Universal Robots URScript: test_fourth_drawing_8_m18.script

def Machining4():
  # Default parameters:
  global speed_ms = 0.3
  global speed_rads = 0.75
  global accel_mss = 3
  global accel_radss = 1.2
  global blend_radius_m = 0.001

  # Add subprograms here
  # Start of main program
  # Program generated by RoboDK v5.6.5 for UR10e on 02/02/2024 17:39:49
  # Using nominal kinematics.
  blend_radius_m = 0.001
  speed_ms = 1.000
  # set_reference(p[0.348734, -0.005000, -0.017586, 0.000000, 0.000000, 0.000000])
  set_tcp(p[0.000000, 0.000000, 0.252000, 0.000000, 0.000000, 0.000000])
  # Show Tool
  movej([0.508484, -0.952512, -2.535391, -1.224486, 1.570796, 2.079280],accel_radss,speed_rads,0,blend_radius_m)
  movel([0.508484, -0.952512, -2.535391, -1.224486, 1.570796, 2.079280],accel_mss,speed_ms,0,blend_radius_m)
  # Splitting Linear movement in 6 (instruction 7: MoveL 3)
  movel([0.508484, -0.969998, -2.560672, -1.181720, 1.570796, 2.079280],accel_mss,speed_ms,0,blend_radius_m)
  movel([0.508484, -0.990214, -2.585461, -1.136714, 1.570796, 2.079280],accel_mss,speed_ms,0,blend_radius_m)
  movel([0.508484, -1.013449, -2.609714, -1.089227, 1.570796, 2.079280],accel_mss,speed_ms,0,blend_radius_m)
  movel([0.508484, -1.040019, -2.633377, -1.038993, 1.570796, 2.079280],accel_mss,speed_ms,0,blend_radius_m)
  movel([0.508484, -1.070270, -2.656387, -0.985731, 1.570796, 2.079280],accel_mss,speed_ms,0,blend_radius_m)
  movel([0.508484, -1.104577, -2.678669, -0.929143, 1.570796, 2.079280],accel_mss,speed_ms,0,blend_radius_m)
  movel([0.508484, -1.104577, -2.678669, -0.929143, 1.570796, 2.079280],accel_mss,speed_ms,0,blend_radius_m)
  speed_ms = 1.000
  movel([0.508484, -1.104577, -2.678669, -0.929143, 1.570796, 2.079280],accel_mss,speed_ms,0,blend_radius_m)
  movel([0.508484, -1.104577, -2.678669, -0.929143, 1.570796, 2.079280],accel_mss,speed_ms,0,blend_radius_m)
  movel([0.508484, -1.104577, -2.678669, -0.929143, 1.570796, 2.079280],accel_mss,speed_ms,0,blend_radius_m)
  speed_ms = 0.005
  movel([0.508484, -1.063908, -2.651841, -0.996640, 1.570796, 2.079280],accel_mss,speed_ms,0,blend_radius_m)
  speed_ms = 1.000
  movel([0.508484, -1.104577, -2.678669, -0.929143, 1.570796, 2.079280],accel_mss,speed_ms,0,blend_radius_m)
  speed_ms = 0.040
  movel([0.508484, -1.104577, -2.678669, -0.929143, 1.570796, 2.079280],accel_mss,speed_ms,0,blend_radius_m)
  speed_ms = 1.000
  movel([0.508484, -1.104577, -2.678669, -0.929143, 1.570796, 2.079280],accel_mss,speed_ms,0,blend_radius_m)
  # Splitting Linear movement in 8 (instruction 21: MoveL 12)
  movel([0.516357, -1.145060, -2.661765, -0.905563, 1.570796, 2.087153],accel_mss,speed_ms,0,blend_radius_m)
  movel([0.523521, -1.183921, -2.644010, -0.884457, 1.570796, 2.094317],accel_mss,speed_ms,0,blend_radius_m)
  movel([0.530064, -1.221217, -2.625467, -0.865705, 1.570796, 2.100861],accel_mss,speed_ms,0,blend_radius_m)
  movel([0.536061, -1.257021, -2.606194, -0.849174, 1.570796, 2.106857],accel_mss,speed_ms,0,blend_radius_m)
  movel([0.541574, -1.291418, -2.586246, -0.834725, 1.570796, 2.112371],accel_mss,speed_ms,0,blend_radius_m)
  movel([0.546659, -1.324498, -2.565672, -0.822220, 1.570796, 2.117455],accel_mss,speed_ms,0,blend_radius_m)
  movel([0.551360, -1.356351, -2.544515, -0.811522, 1.570796, 2.122157],accel_mss,speed_ms,0,blend_radius_m)
  movel([0.555720, -1.387070, -2.522816, -0.802503, 1.570796, 2.126517],accel_mss,speed_ms,0,blend_radius_m)
  speed_ms = 0.005
  movel([0.555720, -1.427952, -2.542321, -0.742116, 1.570796, 2.126517],accel_mss,speed_ms,0,blend_radius_m)
  speed_ms = 0.025
  movel([0.551886, -1.431799, -2.539331, -0.741259, 1.570796, 2.122682],accel_mss,speed_ms,0,blend_radius_m)
  movel([0.549891, -1.433665, -2.537873, -0.740851, 1.570796, 2.120688],accel_mss,speed_ms,0,blend_radius_m)
  movel([0.547837, -1.435468, -2.536459, -0.740462, 1.570796, 2.118634],accel_mss,speed_ms,0,blend_radius_m)
  movel([0.545720, -1.437189, -2.535105, -0.740095, 1.570796, 2.116517],accel_mss,speed_ms,0,blend_radius_m)
  movel([0.543536, -1.438810, -2.533826, -0.739753, 1.570796, 2.114332],accel_mss,speed_ms,0,blend_radius_m)
  movel([0.541277, -1.440313, -2.532636, -0.739441, 1.570796, 2.112073],accel_mss,speed_ms,0,blend_radius_m)
  movel([0.538938, -1.441676, -2.531553, -0.739160, 1.570796, 2.109734],accel_mss,speed_ms,0,blend_radius_m)
  movel([0.539897, -1.440992, -2.532097, -0.739300, 1.570796, 2.110693],accel_mss,speed_ms,0,blend_radius_m)
  movel([0.540974, -1.439974, -2.532904, -0.739511, 1.570796, 2.111771],accel_mss,speed_ms,0,blend_radius_m)
  movel([0.541871, -1.438872, -2.533777, -0.739741, 1.570796, 2.112668],accel_mss,speed_ms,0,blend_radius_m)
  movel([0.542155, -1.438369, -2.534174, -0.739846, 1.570796, 2.112951],accel_mss,speed_ms,0,blend_radius_m)
  movel([0.542280, -1.437941, -2.534512, -0.739936, 1.570796, 2.113076],accel_mss,speed_ms,0,blend_radius_m)
  movel([0.542211, -1.437608, -2.534775, -0.740006, 1.570796, 2.113008],accel_mss,speed_ms,0,blend_radius_m)
  movel([0.541951, -1.437454, -2.534896, -0.740039, 1.570796, 2.112747],accel_mss,speed_ms,0,blend_radius_m)
  movel([0.541528, -1.437461, -2.534891, -0.740037, 1.570796, 2.112324],accel_mss,speed_ms,0,blend_radius_m)
  movel([0.540960, -1.437607, -2.534776, -0.740007, 1.570796, 2.111756],accel_mss,speed_ms,0,blend_radius_m)
  movel([0.539505, -1.438234, -2.534280, -0.739874, 1.570796, 2.110301],accel_mss,speed_ms,0,blend_radius_m)
  movel([0.537786, -1.439172, -2.533539, -0.739678, 1.570796, 2.108582],accel_mss,speed_ms,0,blend_radius_m)
  movel([0.534336, -1.441332, -2.531826, -0.739230, 1.570796, 2.105133],accel_mss,speed_ms,0,blend_radius_m)
  movel([0.532176, -1.442774, -2.530679, -0.738936, 1.570796, 2.102972],accel_mss,speed_ms,0,blend_radius_m)
  movel([0.529059, -1.444697, -2.529144, -0.738548, 1.570796, 2.099855],accel_mss,speed_ms,0,blend_radius_m)
  movel([0.527463, -1.445498, -2.528503, -0.738388, 1.570796, 2.098260],accel_mss,speed_ms,0,blend_radius_m)
  movel([0.525843, -1.446095, -2.528025, -0.738269, 1.570796, 2.096640],accel_mss,speed_ms,0,blend_radius_m)
  movel([0.526257, -1.445821, -2.528245, -0.738324, 1.570796, 2.097053],accel_mss,speed_ms,0,blend_radius_m)
  movel([0.526732, -1.445268, -2.528687, -0.738434, 1.570796, 2.097529],accel_mss,speed_ms,0,blend_radius_m)
  movel([0.527721, -1.443665, -2.529968, -0.738755, 1.570796, 2.098517],accel_mss,speed_ms,0,blend_radius_m)
  movel([0.528500, -1.441980, -2.531312, -0.739098, 1.570796, 2.099296],accel_mss,speed_ms,0,blend_radius_m)
  movel([0.528712, -1.441319, -2.531837, -0.739233, 1.570796, 2.099508],accel_mss,speed_ms,0,blend_radius_m)
  movel([0.528754, -1.440900, -2.532170, -0.739319, 1.570796, 2.099550],accel_mss,speed_ms,0,blend_radius_m)
  movel([0.528518, -1.440358, -2.532599, -0.739431, 1.570796, 2.099315],accel_mss,speed_ms,0,blend_radius_m)
  movel([0.528131, -1.440101, -2.532804, -0.739485, 1.570796, 2.098927],accel_mss,speed_ms,0,blend_radius_m)
  movel([0.527622, -1.440071, -2.532827, -0.739491, 1.570796, 2.098419],accel_mss,speed_ms,0,blend_radius_m)
  movel([0.527024, -1.440220, -2.532709, -0.739460, 1.570796, 2.097821],accel_mss,speed_ms,0,blend_radius_m)
  movel([0.525708, -1.440829, -2.532226, -0.739334, 1.570796, 2.096504],accel_mss,speed_ms,0,blend_radius_m)
  movel([0.524451, -1.441503, -2.531691, -0.739195, 1.570796, 2.095247],accel_mss,speed_ms,0,blend_radius_m)
  movel([0.522478, -1.442423, -2.530959, -0.739007, 1.570796, 2.093274],accel_mss,speed_ms,0,blend_radius_m)
  movel([0.520576, -1.443144, -2.530385, -0.738861, 1.570796, 2.091372],accel_mss,speed_ms,0,blend_radius_m)
  movel([0.518692, -1.443593, -2.530026, -0.738770, 1.570796, 2.089489],accel_mss,speed_ms,0,blend_radius_m)
  movel([0.516787, -1.443689, -2.529949, -0.738750, 1.570796, 2.087583],accel_mss,speed_ms,0,blend_radius_m)
  movel([0.518245, -1.442894, -2.530584, -0.738911, 1.570796, 2.089042],accel_mss,speed_ms,0,blend_radius_m)
  movel([0.519593, -1.441927, -2.531353, -0.739108, 1.570796, 2.090389],accel_mss,speed_ms,0,blend_radius_m)
  movel([0.520169, -1.441329, -2.531829, -0.739231, 1.570796, 2.090965],accel_mss,speed_ms,0,blend_radius_m)
  movel([0.520610, -1.440680, -2.532344, -0.739365, 1.570796, 2.091406],accel_mss,speed_ms,0,blend_radius_m)
  movel([0.520870, -1.440025, -2.532863, -0.739500, 1.570796, 2.091666],accel_mss,speed_ms,0,blend_radius_m)
  movel([0.520888, -1.439417, -2.533345, -0.739627, 1.570796, 2.091684],accel_mss,speed_ms,0,blend_radius_m)
  movel([0.520543, -1.438832, -2.533808, -0.739749, 1.570796, 2.091340],accel_mss,speed_ms,0,blend_radius_m)
  movel([0.519903, -1.438483, -2.534084, -0.739822, 1.570796, 2.090700],accel_mss,speed_ms,0,blend_radius_m)
  movel([0.519080, -1.438310, -2.534221, -0.739858, 1.570796, 2.089876],accel_mss,speed_ms,0,blend_radius_m)
  movel([0.518194, -1.438247, -2.534271, -0.739872, 1.570796, 2.088990],accel_mss,speed_ms,0,blend_radius_m)
  speed_ms = 0.005
  movel([0.518194, -1.429866, -2.530530, -0.751993, 1.570796, 2.088990],accel_mss,speed_ms,0,blend_radius_m)
  speed_ms = 0.040
  movel([0.510141, -1.449455, -2.514970, -0.747963, 1.570796, 2.080938],accel_mss,speed_ms,0,blend_radius_m)
  speed_ms = 0.005
  movel([0.510141, -1.457684, -2.518629, -0.736076, 1.570796, 2.080938],accel_mss,speed_ms,0,blend_radius_m)
  speed_ms = 0.025
  movel([0.511091, -1.456693, -2.519440, -0.736256, 1.570796, 2.081888],accel_mss,speed_ms,0,blend_radius_m)
  movel([0.512141, -1.455770, -2.520195, -0.736424, 1.570796, 2.082937],accel_mss,speed_ms,0,blend_radius_m)
  movel([0.513267, -1.454927, -2.520883, -0.736579, 1.570796, 2.084063],accel_mss,speed_ms,0,blend_radius_m)
  movel([0.514457, -1.454175, -2.521496, -0.736718, 1.570796, 2.085253],accel_mss,speed_ms,0,blend_radius_m)
  movel([0.515692, -1.453521, -2.522028, -0.736840, 1.570796, 2.086488],accel_mss,speed_ms,0,blend_radius_m)
  movel([0.516954, -1.452980, -2.522467, -0.736941, 1.570796, 2.087750],accel_mss,speed_ms,0,blend_radius_m)
  movel([0.518224, -1.452560, -2.522808, -0.737020, 1.570796, 2.089020],accel_mss,speed_ms,0,blend_radius_m)
  movel([0.519487, -1.452271, -2.523043, -0.737075, 1.570796, 2.090284],accel_mss,speed_ms,0,blend_radius_m)
  movel([0.521308, -1.452078, -2.523200, -0.737111, 1.570796, 2.092104],accel_mss,speed_ms,0,blend_radius_m)
  movel([0.522944, -1.452159, -2.523134, -0.737096, 1.570796, 2.093740],accel_mss,speed_ms,0,blend_radius_m)
  movel([0.524404, -1.452488, -2.522867, -0.737034, 1.570796, 2.095200],accel_mss,speed_ms,0,blend_radius_m)
  movel([0.525694, -1.453041, -2.522418, -0.736930, 1.570796, 2.096491],accel_mss,speed_ms,0,blend_radius_m)
  movel([0.526823, -1.453792, -2.521807, -0.736790, 1.570796, 2.097619],accel_mss,speed_ms,0,blend_radius_m)
  movel([0.527798, -1.454719, -2.521052, -0.736618, 1.570796, 2.098594],accel_mss,speed_ms,0,blend_radius_m)
  movel([0.528624, -1.455797, -2.520173, -0.736419, 1.570796, 2.099421],accel_mss,speed_ms,0,blend_radius_m)
  movel([0.529313, -1.457000, -2.519189, -0.736200, 1.570796, 2.100109],accel_mss,speed_ms,0,blend_radius_m)
  movel([0.529870, -1.458305, -2.518119, -0.735965, 1.570796, 2.100667],accel_mss,speed_ms,0,blend_radius_m)
  movel([0.530307, -1.459689, -2.516982, -0.735718, 1.570796, 2.101103],accel_mss,speed_ms,0,blend_radius_m)
  movel([0.530848, -1.462592, -2.514587, -0.735210, 1.570796, 2.101644],accel_mss,speed_ms,0,blend_radius_m)
  movel([0.531006, -1.465517, -2.512160, -0.734712, 1.570796, 2.101803],accel_mss,speed_ms,0,blend_radius_m)
  movel([0.530842, -1.468282, -2.509854, -0.734253, 1.570796, 2.101639],accel_mss,speed_ms,0,blend_radius_m)
  movel([0.530390, -1.471193, -2.507413, -0.733783, 1.570796, 2.101186],accel_mss,speed_ms,0,blend_radius_m)
  movel([0.529720, -1.474131, -2.504936, -0.733322, 1.570796, 2.100516],accel_mss,speed_ms,0,blend_radius_m)
  movel([0.528861, -1.477086, -2.502431, -0.732872, 1.570796, 2.099658],accel_mss,speed_ms,0,blend_radius_m)
  movel([0.527841, -1.480049, -2.499906, -0.732435, 1.570796, 2.098637],accel_mss,speed_ms,0,blend_radius_m)
  movel([0.526687, -1.483008, -2.497369, -0.732012, 1.570796, 2.097483],accel_mss,speed_ms,0,blend_radius_m)
  movel([0.525429, -1.485956, -2.494829, -0.731604, 1.570796, 2.096225],accel_mss,speed_ms,0,blend_radius_m)
  movel([0.522707, -1.491776, -2.489774, -0.730839, 1.570796, 2.093504],accel_mss,speed_ms,0,blend_radius_m)
  movel([0.520789, -1.495817, -2.486233, -0.730340, 1.570796, 2.091586],accel_mss,speed_ms,0,blend_radius_m)
  movel([0.519999, -1.497823, -2.484465, -0.730101, 1.570796, 2.090795],accel_mss,speed_ms,0,blend_radius_m)
  movel([0.519432, -1.499808, -2.482709, -0.729872, 1.570796, 2.090228],accel_mss,speed_ms,0,blend_radius_m)
  movel([0.519026, -1.502378, -2.480427, -0.729584, 1.570796, 2.089822],accel_mss,speed_ms,0,blend_radius_m)
  movel([0.518624, -1.504952, -2.478131, -0.729306, 1.570796, 2.089420],accel_mss,speed_ms,0,blend_radius_m)
  movel([0.518292, -1.506214, -2.477001, -0.729174, 1.570796, 2.089088],accel_mss,speed_ms,0,blend_radius_m)
  movel([0.517800, -1.507448, -2.475895, -0.729047, 1.570796, 2.088596],accel_mss,speed_ms,0,blend_radius_m)
  movel([0.517098, -1.508640, -2.474823, -0.728926, 1.570796, 2.087894],accel_mss,speed_ms,0,blend_radius_m)
  movel([0.516134, -1.509785, -2.473791, -0.728813, 1.570796, 2.086930],accel_mss,speed_ms,0,blend_radius_m)
  movel([0.518755, -1.507097, -2.476210, -0.729083, 1.570796, 2.089552],accel_mss,speed_ms,0,blend_radius_m)
  movel([0.521247, -1.504345, -2.478673, -0.729371, 1.570796, 2.092043],accel_mss,speed_ms,0,blend_radius_m)
  movel([0.526020, -1.498683, -2.483705, -0.730001, 1.570796, 2.096816],accel_mss,speed_ms,0,blend_radius_m)
  movel([0.528599, -1.495468, -2.486539, -0.730382, 1.570796, 2.099395],accel_mss,speed_ms,0,blend_radius_m)
  movel([0.531106, -1.492207, -2.489397, -0.730784, 1.570796, 2.101903],accel_mss,speed_ms,0,blend_radius_m)
  movel([0.535966, -1.485569, -2.495163, -0.731657, 1.570796, 2.106762],accel_mss,speed_ms,0,blend_radius_m)
  movel([0.540563, -1.478943, -2.500850, -0.732596, 1.570796, 2.111359],accel_mss,speed_ms,0,blend_radius_m)
  movel([0.542732, -1.475555, -2.503731, -0.733104, 1.570796, 2.113528],accel_mss,speed_ms,0,blend_radius_m)
  movel([0.544723, -1.472142, -2.506614, -0.733633, 1.570796, 2.115519],accel_mss,speed_ms,0,blend_radius_m)
  movel([0.546112, -1.469422, -2.508900, -0.734068, 1.570796, 2.116908],accel_mss,speed_ms,0,blend_radius_m)
  movel([0.547394, -1.466668, -2.511201, -0.734519, 1.570796, 2.118190],accel_mss,speed_ms,0,blend_radius_m)
  movel([0.548701, -1.463889, -2.513512, -0.734988, 1.570796, 2.119497],accel_mss,speed_ms,0,blend_radius_m)
  movel([0.550164, -1.461093, -2.515825, -0.735471, 1.570796, 2.120961],accel_mss,speed_ms,0,blend_radius_m)
  movel([0.550637, -1.460364, -2.516426, -0.735599, 1.570796, 2.121434],accel_mss,speed_ms,0,blend_radius_m)
  movel([0.551236, -1.459675, -2.516993, -0.735720, 1.570796, 2.122032],accel_mss,speed_ms,0,blend_radius_m)
  movel([0.551916, -1.459170, -2.517409, -0.735810, 1.570796, 2.122713],accel_mss,speed_ms,0,blend_radius_m)
  movel([0.552279, -1.459029, -2.517525, -0.735835, 1.570796, 2.123075],accel_mss,speed_ms,0,blend_radius_m)
  movel([0.552650, -1.458984, -2.517562, -0.735843, 1.570796, 2.123447],accel_mss,speed_ms,0,blend_radius_m)
  movel([0.553094, -1.459095, -2.517470, -0.735823, 1.570796, 2.123890],accel_mss,speed_ms,0,blend_radius_m)
  movel([0.553450, -1.459322, -2.517284, -0.735783, 1.570796, 2.124247],accel_mss,speed_ms,0,blend_radius_m)
  movel([0.555162, -1.460824, -2.516047, -0.735518, 1.570796, 2.125958],accel_mss,speed_ms,0,blend_radius_m)
  movel([0.556530, -1.462499, -2.514664, -0.735226, 1.570796, 2.127326],accel_mss,speed_ms,0,blend_radius_m)
  movel([0.557585, -1.464326, -2.513150, -0.734913, 1.570796, 2.128381],accel_mss,speed_ms,0,blend_radius_m)
  movel([0.558352, -1.466294, -2.511513, -0.734582, 1.570796, 2.129148],accel_mss,speed_ms,0,blend_radius_m)
  movel([0.558858, -1.468380, -2.509772, -0.734237, 1.570796, 2.129655],accel_mss,speed_ms,0,blend_radius_m)
  movel([0.559133, -1.470569, -2.507937, -0.733883, 1.570796, 2.129930],accel_mss,speed_ms,0,blend_radius_m)
  movel([0.559203, -1.472844, -2.506022, -0.733522, 1.570796, 2.129999],accel_mss,speed_ms,0,blend_radius_m)
  movel([0.559091, -1.475191, -2.504039, -0.733159, 1.570796, 2.129888],accel_mss,speed_ms,0,blend_radius_m)
  movel([0.558827, -1.477592, -2.502001, -0.732796, 1.570796, 2.129624],accel_mss,speed_ms,0,blend_radius_m)
  movel([0.558438, -1.480032, -2.499920, -0.732437, 1.570796, 2.129235],accel_mss,speed_ms,0,blend_radius_m)
  movel([0.557386, -1.484964, -2.495685, -0.731739, 1.570796, 2.128183],accel_mss,speed_ms,0,blend_radius_m)
  movel([0.554892, -1.494646, -2.487262, -0.730482, 1.570796, 2.125689],accel_mss,speed_ms,0,blend_radius_m)
  movel([0.554588, -1.496145, -2.485944, -0.730300, 1.570796, 2.125384],accel_mss,speed_ms,0,blend_radius_m)
  movel([0.554575, -1.496851, -2.485322, -0.730216, 1.570796, 2.125371],accel_mss,speed_ms,0,blend_radius_m)
  movel([0.554722, -1.497492, -2.484757, -0.730140, 1.570796, 2.125519],accel_mss,speed_ms,0,blend_radius_m)
  movel([0.555275, -1.498243, -2.484094, -0.730052, 1.570796, 2.126071],accel_mss,speed_ms,0,blend_radius_m)
  movel([0.555655, -1.498482, -2.483883, -0.730024, 1.570796, 2.126451],accel_mss,speed_ms,0,blend_radius_m)
  movel([0.556095, -1.498637, -2.483746, -0.730006, 1.570796, 2.126891],accel_mss,speed_ms,0,blend_radius_m)
  movel([0.557113, -1.498726, -2.483667, -0.729996, 1.570796, 2.127910],accel_mss,speed_ms,0,blend_radius_m)
  movel([0.558266, -1.498560, -2.483813, -0.730015, 1.570796, 2.129063],accel_mss,speed_ms,0,blend_radius_m)
  movel([0.559484, -1.498195, -2.484136, -0.730058, 1.570796, 2.130280],accel_mss,speed_ms,0,blend_radius_m)
  movel([0.560700, -1.497680, -2.484591, -0.730118, 1.570796, 2.131496],accel_mss,speed_ms,0,blend_radius_m)
  movel([0.561849, -1.497066, -2.485132, -0.730190, 1.570796, 2.132646],accel_mss,speed_ms,0,blend_radius_m)
  movel([0.562859, -1.496403, -2.485717, -0.730269, 1.570796, 2.133656],accel_mss,speed_ms,0,blend_radius_m)
  movel([0.564501, -1.495161, -2.486809, -0.730419, 1.570796, 2.135297],accel_mss,speed_ms,0,blend_radius_m)
  movel([0.566103, -1.493854, -2.487956, -0.730579, 1.570796, 2.136900],accel_mss,speed_ms,0,blend_radius_m)
  movel([0.569169, -1.491072, -2.490389, -0.730929, 1.570796, 2.139965],accel_mss,speed_ms,0,blend_radius_m)
  movel([0.572027, -1.488119, -2.492957, -0.731313, 1.570796, 2.142824],accel_mss,speed_ms,0,blend_radius_m)
  movel([0.574646, -1.485054, -2.495608, -0.731727, 1.570796, 2.145443],accel_mss,speed_ms,0,blend_radius_m)
  movel([0.575591, -1.483880, -2.496620, -0.731890, 1.570796, 2.146387],accel_mss,speed_ms,0,blend_radius_m)
  movel([0.576618, -1.482762, -2.497581, -0.732046, 1.570796, 2.147414],accel_mss,speed_ms,0,blend_radius_m)
  movel([0.577188, -1.482268, -2.498005, -0.732116, 1.570796, 2.147985],accel_mss,speed_ms,0,blend_radius_m)
  movel([0.577814, -1.481835, -2.498377, -0.732178, 1.570796, 2.148610],accel_mss,speed_ms,0,blend_radius_m)
  movel([0.578503, -1.481482, -2.498679, -0.732228, 1.570796, 2.149299],accel_mss,speed_ms,0,blend_radius_m)
  movel([0.579266, -1.481229, -2.498896, -0.732264, 1.570796, 2.150062],accel_mss,speed_ms,0,blend_radius_m)
  movel([0.580251, -1.481159, -2.498956, -0.732274, 1.570796, 2.151047],accel_mss,speed_ms,0,blend_radius_m)
  movel([0.581073, -1.481422, -2.498731, -0.732237, 1.570796, 2.151869],accel_mss,speed_ms,0,blend_radius_m)
  movel([0.581707, -1.481932, -2.498293, -0.732164, 1.570796, 2.152503],accel_mss,speed_ms,0,blend_radius_m)
  movel([0.582136, -1.482605, -2.497715, -0.732068, 1.570796, 2.152933],accel_mss,speed_ms,0,blend_radius_m)
  movel([0.582578, -1.483885, -2.496615, -0.731889, 1.570796, 2.153374],accel_mss,speed_ms,0,blend_radius_m)
  movel([0.582850, -1.485265, -2.495426, -0.731698, 1.570796, 2.153646],accel_mss,speed_ms,0,blend_radius_m)
  movel([0.583065, -1.488131, -2.492947, -0.731312, 1.570796, 2.153861],accel_mss,speed_ms,0,blend_radius_m)
  movel([0.583037, -1.489513, -2.491746, -0.731130, 1.570796, 2.153834],accel_mss,speed_ms,0,blend_radius_m)
  movel([0.582882, -1.490891, -2.490546, -0.730952, 1.570796, 2.153679],accel_mss,speed_ms,0,blend_radius_m)
  movel([0.582611, -1.492261, -2.489350, -0.730778, 1.570796, 2.153407],accel_mss,speed_ms,0,blend_radius_m)
  movel([0.582227, -1.493625, -2.488157, -0.730607, 1.570796, 2.153023],accel_mss,speed_ms,0,blend_radius_m)
  movel([0.581738, -1.494980, -2.486969, -0.730441, 1.570796, 2.152535],accel_mss,speed_ms,0,blend_radius_m)
  movel([0.580473, -1.497665, -2.484604, -0.730120, 1.570796, 2.151270],accel_mss,speed_ms,0,blend_radius_m)
  movel([0.579710, -1.498992, -2.483432, -0.729965, 1.570796, 2.150506],accel_mss,speed_ms,0,blend_radius_m)
  movel([0.577960, -1.501613, -2.481108, -0.729668, 1.570796, 2.148756],accel_mss,speed_ms,0,blend_radius_m)
  movel([0.575952, -1.504185, -2.478816, -0.729388, 1.570796, 2.146749],accel_mss,speed_ms,0,blend_radius_m)
  movel([0.573737, -1.506705, -2.476561, -0.729123, 1.570796, 2.144533],accel_mss,speed_ms,0,blend_radius_m)
  movel([0.571371, -1.509163, -2.474352, -0.728874, 1.570796, 2.142167],accel_mss,speed_ms,0,blend_radius_m)
  movel([0.567732, -1.512631, -2.471218, -0.728540, 1.570796, 2.138528],accel_mss,speed_ms,0,blend_radius_m)
  movel([0.565824, -1.514296, -2.469707, -0.728386, 1.570796, 2.136621],accel_mss,speed_ms,0,blend_radius_m)
  movel([0.563854, -1.515893, -2.468253, -0.728243, 1.570796, 2.134651],accel_mss,speed_ms,0,blend_radius_m)
  movel([0.561822, -1.517401, -2.466876, -0.728112, 1.570796, 2.132618],accel_mss,speed_ms,0,blend_radius_m)
  movel([0.559727, -1.518806, -2.465590, -0.727992, 1.570796, 2.130523],accel_mss,speed_ms,0,blend_radius_m)
  movel([0.557561, -1.520091, -2.464412, -0.727886, 1.570796, 2.128357],accel_mss,speed_ms,0,blend_radius_m)
  movel([0.555327, -1.521236, -2.463359, -0.727794, 1.570796, 2.126124],accel_mss,speed_ms,0,blend_radius_m)
  movel([0.552124, -1.522621, -2.462084, -0.727685, 1.570796, 2.122920],accel_mss,speed_ms,0,blend_radius_m)
  movel([0.550419, -1.523230, -2.461521, -0.727638, 1.570796, 2.121215],accel_mss,speed_ms,0,blend_radius_m)
  movel([0.548705, -1.523722, -2.461067, -0.727600, 1.570796, 2.119502],accel_mss,speed_ms,0,blend_radius_m)
  movel([0.547032, -1.524050, -2.460764, -0.727575, 1.570796, 2.117828],accel_mss,speed_ms,0,blend_radius_m)
  movel([0.545444, -1.524166, -2.460656, -0.727567, 1.570796, 2.116240],accel_mss,speed_ms,0,blend_radius_m)
  movel([0.543989, -1.524022, -2.460790, -0.727577, 1.570796, 2.114785],accel_mss,speed_ms,0,blend_radius_m)
  movel([0.543326, -1.523839, -2.460959, -0.727591, 1.570796, 2.114122],accel_mss,speed_ms,0,blend_radius_m)
  movel([0.542715, -1.523572, -2.461206, -0.727611, 1.570796, 2.113512],accel_mss,speed_ms,0,blend_radius_m)
  movel([0.542106, -1.523172, -2.461575, -0.727642, 1.570796, 2.112902],accel_mss,speed_ms,0,blend_radius_m)
  movel([0.541607, -1.522687, -2.462022, -0.727679, 1.570796, 2.112403],accel_mss,speed_ms,0,blend_radius_m)
  movel([0.541207, -1.522126, -2.462540, -0.727723, 1.570796, 2.112004],accel_mss,speed_ms,0,blend_radius_m)
  movel([0.540902, -1.521496, -2.463120, -0.727773, 1.570796, 2.111698],accel_mss,speed_ms,0,blend_radius_m)
  movel([0.540535, -1.520068, -2.464433, -0.727888, 1.570796, 2.111331],accel_mss,speed_ms,0,blend_radius_m)
  movel([0.540444, -1.518473, -2.465896, -0.728020, 1.570796, 2.111240],accel_mss,speed_ms,0,blend_radius_m)
  movel([0.540559, -1.516785, -2.467439, -0.728165, 1.570796, 2.111355],accel_mss,speed_ms,0,blend_radius_m)
  movel([0.540816, -1.515077, -2.468996, -0.728316, 1.570796, 2.111612],accel_mss,speed_ms,0,blend_radius_m)
  movel([0.541487, -1.511892, -2.471888, -0.728610, 1.570796, 2.112284],accel_mss,speed_ms,0,blend_radius_m)
  movel([0.541819, -1.510404, -2.473232, -0.728752, 1.570796, 2.112615],accel_mss,speed_ms,0,blend_radius_m)
  movel([0.541998, -1.508958, -2.474537, -0.728895, 1.570796, 2.112794],accel_mss,speed_ms,0,blend_radius_m)
  movel([0.541952, -1.508290, -2.475137, -0.728961, 1.570796, 2.112748],accel_mss,speed_ms,0,blend_radius_m)
  movel([0.541774, -1.507681, -2.475685, -0.729023, 1.570796, 2.112571],accel_mss,speed_ms,0,blend_radius_m)
  movel([0.541434, -1.507148, -2.476163, -0.729077, 1.570796, 2.112230],accel_mss,speed_ms,0,blend_radius_m)
  movel([0.540901, -1.506706, -2.476560, -0.729123, 1.570796, 2.111697],accel_mss,speed_ms,0,blend_radius_m)
  movel([0.540999, -1.506837, -2.476443, -0.729109, 1.570796, 2.111796],accel_mss,speed_ms,0,blend_radius_m)
  movel([0.540993, -1.507039, -2.476261, -0.729088, 1.570796, 2.111789],accel_mss,speed_ms,0,blend_radius_m)
  movel([0.540687, -1.507637, -2.475725, -0.729027, 1.570796, 2.111483],accel_mss,speed_ms,0,blend_radius_m)
  movel([0.540031, -1.508460, -2.474985, -0.728944, 1.570796, 2.110827],accel_mss,speed_ms,0,blend_radius_m)
  movel([0.539081, -1.509472, -2.474073, -0.728844, 1.570796, 2.109877],accel_mss,speed_ms,0,blend_radius_m)
  movel([0.536506, -1.511911, -2.471870, -0.728608, 1.570796, 2.107302],accel_mss,speed_ms,0,blend_radius_m)
  movel([0.533377, -1.514652, -2.469383, -0.728354, 1.570796, 2.104174],accel_mss,speed_ms,0,blend_radius_m)
  movel([0.527088, -1.519857, -2.464627, -0.727905, 1.570796, 2.097884],accel_mss,speed_ms,0,blend_radius_m)
  movel([0.523408, -1.522733, -2.461980, -0.727676, 1.570796, 2.094204],accel_mss,speed_ms,0,blend_radius_m)
  movel([0.519372, -1.525494, -2.459426, -0.727468, 1.570796, 2.090168],accel_mss,speed_ms,0,blend_radius_m)
  movel([0.515337, -1.528147, -2.456962, -0.727280, 1.570796, 2.086134],accel_mss,speed_ms,0,blend_radius_m)
  movel([0.511276, -1.530728, -2.454553, -0.727108, 1.570796, 2.082072],accel_mss,speed_ms,0,blend_radius_m)
  movel([0.503302, -1.535575, -2.450000, -0.726814, 1.570796, 2.074098],accel_mss,speed_ms,0,blend_radius_m)
  movel([0.499392, -1.537721, -2.447972, -0.726695, 1.570796, 2.070188],accel_mss,speed_ms,0,blend_radius_m)
  movel([0.497416, -1.538674, -2.447070, -0.726645, 1.570796, 2.068213],accel_mss,speed_ms,0,blend_radius_m)
  movel([0.495430, -1.539517, -2.446269, -0.726602, 1.570796, 2.066226],accel_mss,speed_ms,0,blend_radius_m)
  movel([0.493429, -1.540226, -2.445596, -0.726567, 1.570796, 2.064225],accel_mss,speed_ms,0,blend_radius_m)
  movel([0.491417, -1.540779, -2.445070, -0.726540, 1.570796, 2.062214],accel_mss,speed_ms,0,blend_radius_m)
  movel([0.493294, -1.537726, -2.447968, -0.726695, 1.570796, 2.064090],accel_mss,speed_ms,0,blend_radius_m)
  movel([0.493731, -1.536801, -2.448843, -0.726745, 1.570796, 2.064527],accel_mss,speed_ms,0,blend_radius_m)
  movel([0.493771, -1.536384, -2.449237, -0.726768, 1.570796, 2.064567],accel_mss,speed_ms,0,blend_radius_m)
  movel([0.493597, -1.536066, -2.449537, -0.726786, 1.570796, 2.064394],accel_mss,speed_ms,0,blend_radius_m)
  movel([0.493297, -1.535935, -2.449661, -0.726793, 1.570796, 2.064093],accel_mss,speed_ms,0,blend_radius_m)
  movel([0.492915, -1.535922, -2.449673, -0.726794, 1.570796, 2.063711],accel_mss,speed_ms,0,blend_radius_m)
  movel([0.490914, -1.536231, -2.449382, -0.726777, 1.570796, 2.061711],accel_mss,speed_ms,0,blend_radius_m)
  movel([0.489818, -1.536232, -2.449381, -0.726777, 1.570796, 2.060615],accel_mss,speed_ms,0,blend_radius_m)
  movel([0.488797, -1.536075, -2.449529, -0.726785, 1.570796, 2.059594],accel_mss,speed_ms,0,blend_radius_m)
  movel([0.487879, -1.535763, -2.449823, -0.726803, 1.570796, 2.058675],accel_mss,speed_ms,0,blend_radius_m)
  movel([0.487648, -1.535578, -2.449998, -0.726813, 1.570796, 2.058445],accel_mss,speed_ms,0,blend_radius_m)
  movel([0.487677, -1.535333, -2.450228, -0.726827, 1.570796, 2.058473],accel_mss,speed_ms,0,blend_radius_m)
  movel([0.488374, -1.534524, -2.450991, -0.726874, 1.570796, 2.059170],accel_mss,speed_ms,0,blend_radius_m)
  movel([0.488495, -1.534216, -2.451281, -0.726892, 1.570796, 2.059291],accel_mss,speed_ms,0,blend_radius_m)
  movel([0.488458, -1.533935, -2.451545, -0.726909, 1.570796, 2.059254],accel_mss,speed_ms,0,blend_radius_m)
  movel([0.488296, -1.533709, -2.451758, -0.726922, 1.570796, 2.059092],accel_mss,speed_ms,0,blend_radius_m)
  movel([0.488039, -1.533564, -2.451894, -0.726931, 1.570796, 2.058835],accel_mss,speed_ms,0,blend_radius_m)
  movel([0.487372, -1.533509, -2.451945, -0.726934, 1.570796, 2.058169],accel_mss,speed_ms,0,blend_radius_m)
  movel([0.482012, -1.534472, -2.451040, -0.726877, 1.570796, 2.052809],accel_mss,speed_ms,0,blend_radius_m)
  movel([0.483729, -1.533917, -2.451562, -0.726910, 1.570796, 2.054525],accel_mss,speed_ms,0,blend_radius_m)
  movel([0.485480, -1.533241, -2.452198, -0.726951, 1.570796, 2.056276],accel_mss,speed_ms,0,blend_radius_m)
  movel([0.487243, -1.532463, -2.452928, -0.726998, 1.570796, 2.058040],accel_mss,speed_ms,0,blend_radius_m)
  movel([0.489007, -1.531599, -2.453738, -0.727052, 1.570796, 2.059803],accel_mss,speed_ms,0,blend_radius_m)
  movel([0.492467, -1.529679, -2.455534, -0.727177, 1.570796, 2.063264],accel_mss,speed_ms,0,blend_radius_m)
  movel([0.495725, -1.527617, -2.457455, -0.727317, 1.570796, 2.066521],accel_mss,speed_ms,0,blend_radius_m)
  movel([0.499158, -1.525260, -2.459643, -0.727485, 1.570796, 2.069954],accel_mss,speed_ms,0,blend_radius_m)
  movel([0.502533, -1.522773, -2.461943, -0.727673, 1.570796, 2.073330],accel_mss,speed_ms,0,blend_radius_m)
  movel([0.504170, -1.521467, -2.463147, -0.727775, 1.570796, 2.074966],accel_mss,speed_ms,0,blend_radius_m)
  movel([0.505759, -1.520115, -2.464390, -0.727884, 1.570796, 2.076556],accel_mss,speed_ms,0,blend_radius_m)
  movel([0.507286, -1.518712, -2.465677, -0.728000, 1.570796, 2.078082],accel_mss,speed_ms,0,blend_radius_m)
  movel([0.508742, -1.517249, -2.467015, -0.728125, 1.570796, 2.079538],accel_mss,speed_ms,0,blend_radius_m)
  movel([0.509588, -1.516300, -2.467881, -0.728207, 1.570796, 2.080384],accel_mss,speed_ms,0,blend_radius_m)
  movel([0.510366, -1.515308, -2.468786, -0.728295, 1.570796, 2.081163],accel_mss,speed_ms,0,blend_radius_m)
  movel([0.511731, -1.513219, -2.470684, -0.728485, 1.570796, 2.082527],accel_mss,speed_ms,0,blend_radius_m)
  movel([0.512844, -1.511031, -2.472666, -0.728692, 1.570796, 2.083641],accel_mss,speed_ms,0,blend_radius_m)
  movel([0.513716, -1.508789, -2.474689, -0.728912, 1.570796, 2.084513],accel_mss,speed_ms,0,blend_radius_m)
  movel([0.514362, -1.506538, -2.476711, -0.729140, 1.570796, 2.085158],accel_mss,speed_ms,0,blend_radius_m)
  movel([0.514791, -1.504328, -2.478688, -0.729372, 1.570796, 2.085588],accel_mss,speed_ms,0,blend_radius_m)
  movel([0.515013, -1.502206, -2.480580, -0.729603, 1.570796, 2.085809],accel_mss,speed_ms,0,blend_radius_m)
  movel([0.515040, -1.500220, -2.482344, -0.729825, 1.570796, 2.085836],accel_mss,speed_ms,0,blend_radius_m)
  movel([0.514833, -1.499178, -2.483268, -0.729944, 1.570796, 2.085629],accel_mss,speed_ms,0,blend_radius_m)
  movel([0.514328, -1.498388, -2.483965, -0.730035, 1.570796, 2.085125],accel_mss,speed_ms,0,blend_radius_m)
  movel([0.513576, -1.497861, -2.484431, -0.730097, 1.570796, 2.084372],accel_mss,speed_ms,0,blend_radius_m)
  movel([0.512626, -1.497606, -2.484656, -0.730127, 1.570796, 2.083422],accel_mss,speed_ms,0,blend_radius_m)
  movel([0.511527, -1.497627, -2.484638, -0.730124, 1.570796, 2.082323],accel_mss,speed_ms,0,blend_radius_m)
  movel([0.510328, -1.497933, -2.484368, -0.730088, 1.570796, 2.081125],accel_mss,speed_ms,0,blend_radius_m)
  movel([0.509087, -1.498529, -2.483841, -0.730019, 1.570796, 2.079883],accel_mss,speed_ms,0,blend_radius_m)
  movel([0.507849, -1.499420, -2.483053, -0.729916, 1.570796, 2.078646],accel_mss,speed_ms,0,blend_radius_m)
  movel([0.506057, -1.500901, -2.481740, -0.729748, 1.570796, 2.076853],accel_mss,speed_ms,0,blend_radius_m)
  movel([0.504215, -1.502308, -2.480490, -0.729592, 1.570796, 2.075011],accel_mss,speed_ms,0,blend_radius_m)
  movel([0.502327, -1.503615, -2.479325, -0.729449, 1.570796, 2.073123],accel_mss,speed_ms,0,blend_radius_m)
  movel([0.500388, -1.504800, -2.478267, -0.729322, 1.570796, 2.071184],accel_mss,speed_ms,0,blend_radius_m)
  movel([0.498404, -1.505837, -2.477339, -0.729213, 1.570796, 2.069200],accel_mss,speed_ms,0,blend_radius_m)
  movel([0.496371, -1.506704, -2.476562, -0.729123, 1.570796, 2.067167],accel_mss,speed_ms,0,blend_radius_m)
  movel([0.494289, -1.507378, -2.475957, -0.729054, 1.570796, 2.065085],accel_mss,speed_ms,0,blend_radius_m)
  movel([0.492160, -1.507833, -2.475548, -0.729008, 1.570796, 2.062956],accel_mss,speed_ms,0,blend_radius_m)
  movel([0.491077, -1.507930, -2.475462, -0.728998, 1.570796, 2.061873],accel_mss,speed_ms,0,blend_radius_m)
  movel([0.490044, -1.507891, -2.475496, -0.729002, 1.570796, 2.060840],accel_mss,speed_ms,0,blend_radius_m)
  movel([0.488081, -1.507580, -2.475776, -0.729033, 1.570796, 2.058877],accel_mss,speed_ms,0,blend_radius_m)
  movel([0.486632, -1.507175, -2.476139, -0.729075, 1.570796, 2.057428],accel_mss,speed_ms,0,blend_radius_m)
  movel([0.485361, -1.506589, -2.476665, -0.729135, 1.570796, 2.056158],accel_mss,speed_ms,0,blend_radius_m)
  movel([0.484262, -1.505838, -2.477338, -0.729213, 1.570796, 2.055058],accel_mss,speed_ms,0,blend_radius_m)
  movel([0.483321, -1.504938, -2.478144, -0.729308, 1.570796, 2.054117],accel_mss,speed_ms,0,blend_radius_m)
  movel([0.482527, -1.503906, -2.479066, -0.729418, 1.570796, 2.053323],accel_mss,speed_ms,0,blend_radius_m)
  movel([0.481869, -1.502756, -2.480091, -0.729542, 1.570796, 2.052665],accel_mss,speed_ms,0,blend_radius_m)
  movel([0.481342, -1.501504, -2.481204, -0.729680, 1.570796, 2.052138],accel_mss,speed_ms,0,blend_radius_m)
  movel([0.480931, -1.500169, -2.482389, -0.729831, 1.570796, 2.051727],accel_mss,speed_ms,0,blend_radius_m)
  movel([0.480626, -1.498766, -2.483631, -0.729991, 1.570796, 2.051422],accel_mss,speed_ms,0,blend_radius_m)
  movel([0.480420, -1.497308, -2.484919, -0.730162, 1.570796, 2.051216],accel_mss,speed_ms,0,blend_radius_m)
  movel([0.480258, -1.494306, -2.487560, -0.730523, 1.570796, 2.051054],accel_mss,speed_ms,0,blend_radius_m)
  movel([0.480362, -1.491291, -2.490197, -0.730901, 1.570796, 2.051158],accel_mss,speed_ms,0,blend_radius_m)
  movel([0.480649, -1.488405, -2.492708, -0.731275, 1.570796, 2.051445],accel_mss,speed_ms,0,blend_radius_m)
  movel([0.480991, -1.486173, -2.494642, -0.731574, 1.570796, 2.051788],accel_mss,speed_ms,0,blend_radius_m)
  movel([0.481470, -1.483852, -2.496643, -0.731893, 1.570796, 2.052266],accel_mss,speed_ms,0,blend_radius_m)
  movel([0.482087, -1.481456, -2.498701, -0.732232, 1.570796, 2.052883],accel_mss,speed_ms,0,blend_radius_m)
  movel([0.482851, -1.479008, -2.500794, -0.732587, 1.570796, 2.053648],accel_mss,speed_ms,0,blend_radius_m)
  movel([0.483763, -1.476523, -2.502909, -0.732957, 1.570796, 2.054560],accel_mss,speed_ms,0,blend_radius_m)
  movel([0.484830, -1.474022, -2.505028, -0.733339, 1.570796, 2.055627],accel_mss,speed_ms,0,blend_radius_m)
  movel([0.486057, -1.471525, -2.507134, -0.733730, 1.570796, 2.056854],accel_mss,speed_ms,0,blend_radius_m)
  movel([0.487449, -1.469050, -2.509211, -0.734128, 1.570796, 2.058245],accel_mss,speed_ms,0,blend_radius_m)
  movel([0.489008, -1.466616, -2.511245, -0.734528, 1.570796, 2.059805],accel_mss,speed_ms,0,blend_radius_m)
  movel([0.490739, -1.464248, -2.513215, -0.734927, 1.570796, 2.061535],accel_mss,speed_ms,0,blend_radius_m)
  movel([0.492647, -1.461961, -2.515109, -0.735320, 1.570796, 2.063443],accel_mss,speed_ms,0,blend_radius_m)
  movel([0.494736, -1.459780, -2.516907, -0.735702, 1.570796, 2.065532],accel_mss,speed_ms,0,blend_radius_m)
  movel([0.497007, -1.457726, -2.518594, -0.736069, 1.570796, 2.067803],accel_mss,speed_ms,0,blend_radius_m)
  movel([0.499467, -1.455820, -2.520154, -0.736415, 1.570796, 2.070264],accel_mss,speed_ms,0,blend_radius_m)
  movel([0.502114, -1.454087, -2.521567, -0.736735, 1.570796, 2.072911],accel_mss,speed_ms,0,blend_radius_m)
  movel([0.504952, -1.452548, -2.522818, -0.737023, 1.570796, 2.075748],accel_mss,speed_ms,0,blend_radius_m)
  movel([0.506085, -1.452062, -2.523213, -0.737114, 1.570796, 2.076882],accel_mss,speed_ms,0,blend_radius_m)
  movel([0.506646, -1.451910, -2.523336, -0.737143, 1.570796, 2.077442],accel_mss,speed_ms,0,blend_radius_m)
  movel([0.507180, -1.451865, -2.523372, -0.737151, 1.570796, 2.077976],accel_mss,speed_ms,0,blend_radius_m)
  movel([0.507850, -1.452048, -2.523224, -0.737117, 1.570796, 2.078646],accel_mss,speed_ms,0,blend_radius_m)
  movel([0.508305, -1.452476, -2.522877, -0.737036, 1.570796, 2.079101],accel_mss,speed_ms,0,blend_radius_m)
  movel([0.508559, -1.453073, -2.522392, -0.736924, 1.570796, 2.079355],accel_mss,speed_ms,0,blend_radius_m)
  movel([0.508624, -1.453762, -2.521832, -0.736795, 1.570796, 2.079421],accel_mss,speed_ms,0,blend_radius_m)
  movel([0.508371, -1.455391, -2.520505, -0.736494, 1.570796, 2.079167],accel_mss,speed_ms,0,blend_radius_m)
  movel([0.507807, -1.457086, -2.519119, -0.736184, 1.570796, 2.078604],accel_mss,speed_ms,0,blend_radius_m)
  movel([0.506383, -1.460472, -2.516337, -0.735580, 1.570796, 2.077180],accel_mss,speed_ms,0,blend_radius_m)
  movel([0.506259, -1.461115, -2.515807, -0.735467, 1.570796, 2.077056],accel_mss,speed_ms,0,blend_radius_m)
  movel([0.506393, -1.461311, -2.515645, -0.735433, 1.570796, 2.077189],accel_mss,speed_ms,0,blend_radius_m)
  movel([0.506705, -1.461409, -2.515565, -0.735416, 1.570796, 2.077502],accel_mss,speed_ms,0,blend_radius_m)
  movel([0.507835, -1.460385, -2.516409, -0.735595, 1.570796, 2.078631],accel_mss,speed_ms,0,blend_radius_m)
  movel([0.508922, -1.459289, -2.517311, -0.735789, 1.570796, 2.079718],accel_mss,speed_ms,0,blend_radius_m)
  movel([0.506690, -1.464208, -2.513247, -0.734933, 1.570796, 2.077486],accel_mss,speed_ms,0,blend_radius_m)
  movel([0.504647, -1.469094, -2.509174, -0.734121, 1.570796, 2.075443],accel_mss,speed_ms,0,blend_radius_m)
  movel([0.502794, -1.473940, -2.505097, -0.733352, 1.570796, 2.073591],accel_mss,speed_ms,0,blend_radius_m)
  movel([0.501130, -1.478747, -2.501017, -0.732625, 1.570796, 2.071926],accel_mss,speed_ms,0,blend_radius_m)
  movel([0.500482, -1.480827, -2.499240, -0.732322, 1.570796, 2.071279],accel_mss,speed_ms,0,blend_radius_m)
  movel([0.499986, -1.482980, -2.497394, -0.732016, 1.570796, 2.070782],accel_mss,speed_ms,0,blend_radius_m)
  movel([0.499855, -1.484030, -2.496490, -0.731869, 1.570796, 2.070651],accel_mss,speed_ms,0,blend_radius_m)
  movel([0.499835, -1.485034, -2.495625, -0.731730, 1.570796, 2.070632],accel_mss,speed_ms,0,blend_radius_m)
  movel([0.499953, -1.485969, -2.494818, -0.731602, 1.570796, 2.070750],accel_mss,speed_ms,0,blend_radius_m)
  movel([0.500234, -1.486813, -2.494088, -0.731488, 1.570796, 2.071030],accel_mss,speed_ms,0,blend_radius_m)
  movel([0.500540, -1.487327, -2.493643, -0.731419, 1.570796, 2.071337],accel_mss,speed_ms,0,blend_radius_m)
  movel([0.501409, -1.488098, -2.492975, -0.731316, 1.570796, 2.072205],accel_mss,speed_ms,0,blend_radius_m)
  movel([0.501954, -1.488363, -2.492745, -0.731281, 1.570796, 2.072751],accel_mss,speed_ms,0,blend_radius_m)
  movel([0.503221, -1.488682, -2.492468, -0.731239, 1.570796, 2.074017],accel_mss,speed_ms,0,blend_radius_m)
  movel([0.504669, -1.488745, -2.492413, -0.731231, 1.570796, 2.075466],accel_mss,speed_ms,0,blend_radius_m)
  movel([0.506229, -1.488592, -2.492546, -0.731251, 1.570796, 2.077025],accel_mss,speed_ms,0,blend_radius_m)
  movel([0.507834, -1.488256, -2.492838, -0.731295, 1.570796, 2.078630],accel_mss,speed_ms,0,blend_radius_m)
  movel([0.509415, -1.487776, -2.493254, -0.731359, 1.570796, 2.080211],accel_mss,speed_ms,0,blend_radius_m)
  movel([0.510902, -1.487184, -2.493767, -0.731438, 1.570796, 2.081698],accel_mss,speed_ms,0,blend_radius_m)
  speed_ms = 0.005
  movel([0.510902, -1.479192, -2.490228, -0.742968, 1.570796, 2.081698],accel_mss,speed_ms,0,blend_radius_m)
  speed_ms = 0.040
  movel([0.504315, -1.478811, -2.490555, -0.743024, 1.570796, 2.075111],accel_mss,speed_ms,0,blend_radius_m)
  speed_ms = 0.005
  movel([0.504315, -1.486806, -2.494094, -0.731489, 1.570796, 2.075111],accel_mss,speed_ms,0,blend_radius_m)
  speed_ms = 0.025
  movel([0.505537, -1.486277, -2.494552, -0.731560, 1.570796, 2.076334],accel_mss,speed_ms,0,blend_radius_m)
  movel([0.508048, -1.484927, -2.495717, -0.731745, 1.570796, 2.078844],accel_mss,speed_ms,0,blend_radius_m)
  movel([0.509310, -1.484124, -2.496410, -0.731856, 1.570796, 2.080107],accel_mss,speed_ms,0,blend_radius_m)
  movel([0.511786, -1.482304, -2.497974, -0.732111, 1.570796, 2.082582],accel_mss,speed_ms,0,blend_radius_m)
  movel([0.514121, -1.480259, -2.499726, -0.732404, 1.570796, 2.084918],accel_mss,speed_ms,0,blend_radius_m)
  movel([0.515205, -1.479174, -2.500652, -0.732562, 1.570796, 2.086001],accel_mss,speed_ms,0,blend_radius_m)
  movel([0.516215, -1.478057, -2.501605, -0.732727, 1.570796, 2.087012],accel_mss,speed_ms,0,blend_radius_m)
  movel([0.517967, -1.475769, -2.503549, -0.733071, 1.570796, 2.088763],accel_mss,speed_ms,0,blend_radius_m)
  movel([0.518685, -1.474614, -2.504528, -0.733248, 1.570796, 2.089481],accel_mss,speed_ms,0,blend_radius_m)
  movel([0.519277, -1.473465, -2.505498, -0.733425, 1.570796, 2.090073],accel_mss,speed_ms,0,blend_radius_m)
  movel([0.519733, -1.472331, -2.506455, -0.733603, 1.570796, 2.090530],accel_mss,speed_ms,0,blend_radius_m)
  movel([0.520040, -1.471221, -2.507390, -0.733779, 1.570796, 2.090837],accel_mss,speed_ms,0,blend_radius_m)
  movel([0.520253, -1.469872, -2.508522, -0.733995, 1.570796, 2.091049],accel_mss,speed_ms,0,blend_radius_m)
  movel([0.520313, -1.468570, -2.509613, -0.734206, 1.570796, 2.091109],accel_mss,speed_ms,0,blend_radius_m)
  movel([0.520194, -1.467346, -2.510636, -0.734407, 1.570796, 2.090990],accel_mss,speed_ms,0,blend_radius_m)
  movel([0.519870, -1.466239, -2.511559, -0.734591, 1.570796, 2.090666],accel_mss,speed_ms,0,blend_radius_m)
  movel([0.519315, -1.465282, -2.512355, -0.734751, 1.570796, 2.090111],accel_mss,speed_ms,0,blend_radius_m)
  movel([0.518505, -1.464514, -2.512994, -0.734881, 1.570796, 2.089301],accel_mss,speed_ms,0,blend_radius_m)
  movel([0.517413, -1.463971, -2.513444, -0.734974, 1.570796, 2.088209],accel_mss,speed_ms,0,blend_radius_m)
  movel([0.516017, -1.463685, -2.513681, -0.735023, 1.570796, 2.086813],accel_mss,speed_ms,0,blend_radius_m)
  movel([0.514950, -1.463686, -2.513680, -0.735022, 1.570796, 2.085747],accel_mss,speed_ms,0,blend_radius_m)
  movel([0.513820, -1.463866, -2.513531, -0.734992, 1.570796, 2.084616],accel_mss,speed_ms,0,blend_radius_m)
  movel([0.512668, -1.464211, -2.513245, -0.734933, 1.570796, 2.083464],accel_mss,speed_ms,0,blend_radius_m)
  movel([0.511531, -1.464705, -2.512835, -0.734849, 1.570796, 2.082327],accel_mss,speed_ms,0,blend_radius_m)
  movel([0.510447, -1.465335, -2.512311, -0.734743, 1.570796, 2.081243],accel_mss,speed_ms,0,blend_radius_m)
  movel([0.509455, -1.466086, -2.511687, -0.734617, 1.570796, 2.080251],accel_mss,speed_ms,0,blend_radius_m)
  movel([0.508594, -1.466942, -2.510973, -0.734474, 1.570796, 2.079391],accel_mss,speed_ms,0,blend_radius_m)
  movel([0.507900, -1.467889, -2.510182, -0.734318, 1.570796, 2.078696],accel_mss,speed_ms,0,blend_radius_m)
  speed_ms = 0.005
  movel([0.507900, -1.459742, -2.506566, -0.746082, 1.570796, 2.078696],accel_mss,speed_ms,0,blend_radius_m)
  speed_ms = 0.040
  # Splitting Linear movement in 2 (instruction 399: MoveL 378)
  movel([0.523348, -1.483026, -2.486939, -0.742424, 1.570796, 2.094144],accel_mss,speed_ms,0,blend_radius_m)
  movel([0.537863, -1.506106, -2.466651, -0.739632, 1.570796, 2.108659],accel_mss,speed_ms,0,blend_radius_m)
  speed_ms = 0.005
  movel([0.537863, -1.513881, -2.470084, -0.728424, 1.570796, 2.108659],accel_mss,speed_ms,0,blend_radius_m)
  speed_ms = 0.025
  movel([0.534804, -1.518746, -2.465646, -0.727997, 1.570796, 2.105600],accel_mss,speed_ms,0,blend_radius_m)
  movel([0.533121, -1.521109, -2.463476, -0.727804, 1.570796, 2.103918],accel_mss,speed_ms,0,blend_radius_m)
  movel([0.532179, -1.522267, -2.462410, -0.727712, 1.570796, 2.102975],accel_mss,speed_ms,0,blend_radius_m)
  movel([0.531146, -1.523403, -2.461362, -0.727624, 1.570796, 2.101942],accel_mss,speed_ms,0,blend_radius_m)
  movel([0.529945, -1.524547, -2.460304, -0.727538, 1.570796, 2.100741],accel_mss,speed_ms,0,blend_radius_m)
  movel([0.529289, -1.525058, -2.459830, -0.727500, 1.570796, 2.100085],accel_mss,speed_ms,0,blend_radius_m)
  movel([0.528582, -1.525499, -2.459422, -0.727468, 1.570796, 2.099378],accel_mss,speed_ms,0,blend_radius_m)
  movel([0.529133, -1.524304, -2.460528, -0.727556, 1.570796, 2.099929],accel_mss,speed_ms,0,blend_radius_m)
  movel([0.529482, -1.523112, -2.461630, -0.727647, 1.570796, 2.100279],accel_mss,speed_ms,0,blend_radius_m)
  movel([0.529474, -1.522730, -2.461983, -0.727676, 1.570796, 2.100270],accel_mss,speed_ms,0,blend_radius_m)
  movel([0.529326, -1.522627, -2.462078, -0.727684, 1.570796, 2.100123],accel_mss,speed_ms,0,blend_radius_m)
  movel([0.529110, -1.522609, -2.462095, -0.727685, 1.570796, 2.099906],accel_mss,speed_ms,0,blend_radius_m)
  movel([0.528595, -1.522751, -2.461963, -0.727674, 1.570796, 2.099391],accel_mss,speed_ms,0,blend_radius_m)
  movel([0.527773, -1.523173, -2.461574, -0.727642, 1.570796, 2.098570],accel_mss,speed_ms,0,blend_radius_m)
  movel([0.527042, -1.523682, -2.461104, -0.727603, 1.570796, 2.097839],accel_mss,speed_ms,0,blend_radius_m)
  movel([0.526387, -1.524259, -2.460570, -0.727560, 1.570796, 2.097183],accel_mss,speed_ms,0,blend_radius_m)
  movel([0.525792, -1.524887, -2.459990, -0.727513, 1.570796, 2.096588],accel_mss,speed_ms,0,blend_radius_m)
  movel([0.523657, -1.527569, -2.457500, -0.727320, 1.570796, 2.094453],accel_mss,speed_ms,0,blend_radius_m)
  movel([0.522328, -1.529102, -2.456072, -0.727215, 1.570796, 2.093124],accel_mss,speed_ms,0,blend_radius_m)
  movel([0.520904, -1.530578, -2.454693, -0.727118, 1.570796, 2.091700],accel_mss,speed_ms,0,blend_radius_m)
  movel([0.519366, -1.531969, -2.453391, -0.727029, 1.570796, 2.090162],accel_mss,speed_ms,0,blend_radius_m)
  movel([0.517701, -1.533238, -2.452200, -0.726951, 1.570796, 2.088497],accel_mss,speed_ms,0,blend_radius_m)
  movel([0.518592, -1.531972, -2.453389, -0.727029, 1.570796, 2.089388],accel_mss,speed_ms,0,blend_radius_m)
  movel([0.519175, -1.530653, -2.454623, -0.727113, 1.570796, 2.089972],accel_mss,speed_ms,0,blend_radius_m)
  movel([0.519249, -1.530320, -2.454934, -0.727134, 1.570796, 2.090045],accel_mss,speed_ms,0,blend_radius_m)
  movel([0.519182, -1.530039, -2.455197, -0.727153, 1.570796, 2.089978],accel_mss,speed_ms,0,blend_radius_m)
  movel([0.518981, -1.529919, -2.455309, -0.727161, 1.570796, 2.089777],accel_mss,speed_ms,0,blend_radius_m)
  movel([0.518695, -1.529909, -2.455318, -0.727161, 1.570796, 2.089492],accel_mss,speed_ms,0,blend_radius_m)
  movel([0.518041, -1.530107, -2.455134, -0.727148, 1.570796, 2.088838],accel_mss,speed_ms,0,blend_radius_m)
  movel([0.517247, -1.530525, -2.454743, -0.727121, 1.570796, 2.088044],accel_mss,speed_ms,0,blend_radius_m)
  movel([0.516500, -1.531034, -2.454266, -0.727088, 1.570796, 2.087296],accel_mss,speed_ms,0,blend_radius_m)
  movel([0.515121, -1.532230, -2.453147, -0.727013, 1.570796, 2.085917],accel_mss,speed_ms,0,blend_radius_m)
  movel([0.512588, -1.534774, -2.450755, -0.726860, 1.570796, 2.083384],accel_mss,speed_ms,0,blend_radius_m)
  movel([0.511075, -1.536112, -2.449494, -0.726783, 1.570796, 2.081871],accel_mss,speed_ms,0,blend_radius_m)
  movel([0.509482, -1.537370, -2.448304, -0.726714, 1.570796, 2.080278],accel_mss,speed_ms,0,blend_radius_m)
  movel([0.507801, -1.538507, -2.447228, -0.726654, 1.570796, 2.078597],accel_mss,speed_ms,0,blend_radius_m)
  movel([0.506025, -1.539481, -2.446304, -0.726604, 1.570796, 2.076821],accel_mss,speed_ms,0,blend_radius_m)
  movel([0.506593, -1.538824, -2.446928, -0.726638, 1.570796, 2.077389],accel_mss,speed_ms,0,blend_radius_m)
  movel([0.507483, -1.537432, -2.448246, -0.726711, 1.570796, 2.078279],accel_mss,speed_ms,0,blend_radius_m)
  movel([0.507792, -1.536717, -2.448922, -0.726750, 1.570796, 2.078589],accel_mss,speed_ms,0,blend_radius_m)
  movel([0.507859, -1.536388, -2.449233, -0.726768, 1.570796, 2.078655],accel_mss,speed_ms,0,blend_radius_m)
  movel([0.507713, -1.536176, -2.449433, -0.726780, 1.570796, 2.078509],accel_mss,speed_ms,0,blend_radius_m)
  movel([0.507336, -1.536230, -2.449382, -0.726777, 1.570796, 2.078132],accel_mss,speed_ms,0,blend_radius_m)
  movel([0.506369, -1.536616, -2.449017, -0.726755, 1.570796, 2.077165],accel_mss,speed_ms,0,blend_radius_m)
  movel([0.505468, -1.537086, -2.448573, -0.726730, 1.570796, 2.076264],accel_mss,speed_ms,0,blend_radius_m)
  movel([0.503783, -1.538190, -2.447528, -0.726671, 1.570796, 2.074579],accel_mss,speed_ms,0,blend_radius_m)
  movel([0.502119, -1.539347, -2.446431, -0.726611, 1.570796, 2.072916],accel_mss,speed_ms,0,blend_radius_m)
  movel([0.501243, -1.539886, -2.445919, -0.726584, 1.570796, 2.072040],accel_mss,speed_ms,0,blend_radius_m)
  movel([0.500309, -1.540369, -2.445461, -0.726560, 1.570796, 2.071105],accel_mss,speed_ms,0,blend_radius_m)
  movel([0.497992, -1.541360, -2.444518, -0.726512, 1.570796, 2.068789],accel_mss,speed_ms,0,blend_radius_m)
  movel([0.495656, -1.542234, -2.443684, -0.726471, 1.570796, 2.066453],accel_mss,speed_ms,0,blend_radius_m)
  movel([0.493314, -1.543007, -2.442947, -0.726436, 1.570796, 2.064111],accel_mss,speed_ms,0,blend_radius_m)
  movel([0.490972, -1.543698, -2.442286, -0.726405, 1.570796, 2.061768],accel_mss,speed_ms,0,blend_radius_m)
  speed_ms = 0.005
  movel([0.490972, -1.536166, -2.438968, -0.737255, 1.570796, 2.061768],accel_mss,speed_ms,0,blend_radius_m)
  speed_ms = 0.040
  movel([0.487780, -1.510169, -2.462992, -0.739227, 1.570796, 2.058576],accel_mss,speed_ms,0,blend_radius_m)
  speed_ms = 0.005
  movel([0.487780, -1.517912, -2.466409, -0.728068, 1.570796, 2.058576],accel_mss,speed_ms,0,blend_radius_m)
  speed_ms = 0.025
  movel([0.488572, -1.517575, -2.466717, -0.728097, 1.570796, 2.059368],accel_mss,speed_ms,0,blend_radius_m)
  movel([0.489350, -1.517128, -2.467126, -0.728135, 1.570796, 2.060146],accel_mss,speed_ms,0,blend_radius_m)
  movel([0.490888, -1.516039, -2.468120, -0.728230, 1.570796, 2.061684],accel_mss,speed_ms,0,blend_radius_m)
  movel([0.492434, -1.514904, -2.469154, -0.728331, 1.570796, 2.063230],accel_mss,speed_ms,0,blend_radius_m)
  movel([0.493224, -1.514400, -2.469612, -0.728377, 1.570796, 2.064021],accel_mss,speed_ms,0,blend_radius_m)
  movel([0.494032, -1.513985, -2.469990, -0.728415, 1.570796, 2.064828],accel_mss,speed_ms,0,blend_radius_m)
  movel([0.494623, -1.513764, -2.470190, -0.728435, 1.570796, 2.065419],accel_mss,speed_ms,0,blend_radius_m)
  movel([0.495063, -1.513684, -2.470262, -0.728442, 1.570796, 2.065860],accel_mss,speed_ms,0,blend_radius_m)
  movel([0.495369, -1.513727, -2.470223, -0.728438, 1.570796, 2.066165],accel_mss,speed_ms,0,blend_radius_m)
  movel([0.495556, -1.513878, -2.470087, -0.728425, 1.570796, 2.066352],accel_mss,speed_ms,0,blend_radius_m)
  movel([0.495622, -1.514444, -2.469572, -0.728373, 1.570796, 2.066419],accel_mss,speed_ms,0,blend_radius_m)
  movel([0.495380, -1.515256, -2.468833, -0.728300, 1.570796, 2.066176],accel_mss,speed_ms,0,blend_radius_m)
  movel([0.494420, -1.517121, -2.467132, -0.728136, 1.570796, 2.065216],accel_mss,speed_ms,0,blend_radius_m)
  movel([0.493590, -1.518486, -2.465884, -0.728019, 1.570796, 2.064386],accel_mss,speed_ms,0,blend_radius_m)
  movel([0.495203, -1.517431, -2.466849, -0.728109, 1.570796, 2.065999],accel_mss,speed_ms,0,blend_radius_m)
  movel([0.496592, -1.516279, -2.467900, -0.728209, 1.570796, 2.067388],accel_mss,speed_ms,0,blend_radius_m)
  movel([0.497820, -1.515050, -2.469020, -0.728318, 1.570796, 2.068616],accel_mss,speed_ms,0,blend_radius_m)
  movel([0.498939, -1.513767, -2.470188, -0.728435, 1.570796, 2.069735],accel_mss,speed_ms,0,blend_radius_m)
  movel([0.502214, -1.509791, -2.473786, -0.728812, 1.570796, 2.073011],accel_mss,speed_ms,0,blend_radius_m)
  movel([0.503467, -1.508496, -2.474952, -0.728941, 1.570796, 2.074264],accel_mss,speed_ms,0,blend_radius_m)
  movel([0.504042, -1.508033, -2.475369, -0.728987, 1.570796, 2.074839],accel_mss,speed_ms,0,blend_radius_m)
  movel([0.504505, -1.507825, -2.475555, -0.729008, 1.570796, 2.075301],accel_mss,speed_ms,0,blend_radius_m)
  movel([0.504864, -1.507828, -2.475553, -0.729008, 1.570796, 2.075660],accel_mss,speed_ms,0,blend_radius_m)
  movel([0.505123, -1.508000, -2.475398, -0.728991, 1.570796, 2.075919],accel_mss,speed_ms,0,blend_radius_m)
  movel([0.505294, -1.508296, -2.475132, -0.728961, 1.570796, 2.076091],accel_mss,speed_ms,0,blend_radius_m)
  movel([0.505381, -1.508672, -2.474794, -0.728923, 1.570796, 2.076177],accel_mss,speed_ms,0,blend_radius_m)
  movel([0.505338, -1.509493, -2.474054, -0.728842, 1.570796, 2.076134],accel_mss,speed_ms,0,blend_radius_m)
  movel([0.505014, -1.510325, -2.473304, -0.728760, 1.570796, 2.075810],accel_mss,speed_ms,0,blend_radius_m)
  movel([0.504439, -1.511358, -2.472370, -0.728660, 1.570796, 2.075235],accel_mss,speed_ms,0,blend_radius_m)
  movel([0.503263, -1.513232, -2.470673, -0.728484, 1.570796, 2.074059],accel_mss,speed_ms,0,blend_radius_m)
  movel([0.505626, -1.510620, -2.473038, -0.728732, 1.570796, 2.076422],accel_mss,speed_ms,0,blend_radius_m)
  movel([0.506698, -1.509260, -2.474264, -0.728865, 1.570796, 2.077494],accel_mss,speed_ms,0,blend_radius_m)
  movel([0.508605, -1.506453, -2.476787, -0.729149, 1.570796, 2.079402],accel_mss,speed_ms,0,blend_radius_m)
  movel([0.509431, -1.505018, -2.478072, -0.729299, 1.570796, 2.080227],accel_mss,speed_ms,0,blend_radius_m)
  movel([0.510811, -1.502110, -2.480666, -0.729613, 1.570796, 2.081607],accel_mss,speed_ms,0,blend_radius_m)
  speed_ms = 0.005
  movel([0.510811, -1.494239, -2.477187, -0.740963, 1.570796, 2.081607],accel_mss,speed_ms,0,blend_radius_m)
  speed_ms = 0.040
  movel([0.497117, -1.501666, -2.470618, -0.740104, 1.570796, 2.067913],accel_mss,speed_ms,0,blend_radius_m)
  speed_ms = 0.005
  movel([0.497117, -1.509478, -2.474068, -0.728843, 1.570796, 2.067913],accel_mss,speed_ms,0,blend_radius_m)
  speed_ms = 0.025
  movel([0.495257, -1.510649, -2.473012, -0.728729, 1.570796, 2.066053],accel_mss,speed_ms,0,blend_radius_m)
  movel([0.493461, -1.511915, -2.471867, -0.728607, 1.570796, 2.064257],accel_mss,speed_ms,0,blend_radius_m)
  movel([0.489912, -1.514496, -2.469525, -0.728368, 1.570796, 2.060708],accel_mss,speed_ms,0,blend_radius_m)
  movel([0.488066, -1.515701, -2.468428, -0.728260, 1.570796, 2.058863],accel_mss,speed_ms,0,blend_radius_m)
  movel([0.486153, -1.516758, -2.467464, -0.728167, 1.570796, 2.056949],accel_mss,speed_ms,0,blend_radius_m)
  movel([0.484199, -1.517579, -2.466714, -0.728096, 1.570796, 2.054996],accel_mss,speed_ms,0,blend_radius_m)
  movel([0.483218, -1.517873, -2.466445, -0.728071, 1.570796, 2.054014],accel_mss,speed_ms,0,blend_radius_m)
  movel([0.482238, -1.518076, -2.466259, -0.728054, 1.570796, 2.053034],accel_mss,speed_ms,0,blend_radius_m)
  movel([0.483018, -1.517797, -2.466514, -0.728078, 1.570796, 2.053815],accel_mss,speed_ms,0,blend_radius_m)
  movel([0.483969, -1.517228, -2.467035, -0.728127, 1.570796, 2.054765],accel_mss,speed_ms,0,blend_radius_m)
  movel([0.484967, -1.516459, -2.467736, -0.728193, 1.570796, 2.055763],accel_mss,speed_ms,0,blend_radius_m)
  movel([0.485881, -1.515585, -2.468533, -0.728270, 1.570796, 2.056677],accel_mss,speed_ms,0,blend_radius_m)
  movel([0.486585, -1.514696, -2.469343, -0.728350, 1.570796, 2.057381],accel_mss,speed_ms,0,blend_radius_m)
  movel([0.486814, -1.514276, -2.469725, -0.728388, 1.570796, 2.057611],accel_mss,speed_ms,0,blend_radius_m)
  movel([0.486945, -1.513888, -2.470078, -0.728424, 1.570796, 2.057741],accel_mss,speed_ms,0,blend_radius_m)
  movel([0.486958, -1.513541, -2.470392, -0.728455, 1.570796, 2.057755],accel_mss,speed_ms,0,blend_radius_m)
  movel([0.486836, -1.513251, -2.470656, -0.728482, 1.570796, 2.057632],accel_mss,speed_ms,0,blend_radius_m)
  movel([0.486566, -1.513027, -2.470859, -0.728503, 1.570796, 2.057362],accel_mss,speed_ms,0,blend_radius_m)
  movel([0.486127, -1.512881, -2.470991, -0.728517, 1.570796, 2.056923],accel_mss,speed_ms,0,blend_radius_m)
  movel([0.485294, -1.512904, -2.470970, -0.728514, 1.570796, 2.056090],accel_mss,speed_ms,0,blend_radius_m)
  movel([0.481486, -1.513751, -2.470201, -0.728436, 1.570796, 2.052282],accel_mss,speed_ms,0,blend_radius_m)
  movel([0.479925, -1.513965, -2.470008, -0.728417, 1.570796, 2.050722],accel_mss,speed_ms,0,blend_radius_m)
  movel([0.478382, -1.514060, -2.469921, -0.728408, 1.570796, 2.049179],accel_mss,speed_ms,0,blend_radius_m)
  movel([0.476919, -1.514007, -2.469969, -0.728413, 1.570796, 2.047715],accel_mss,speed_ms,0,blend_radius_m)
  movel([0.475600, -1.513769, -2.470186, -0.728435, 1.570796, 2.046397],accel_mss,speed_ms,0,blend_radius_m)
  movel([0.474488, -1.513312, -2.470600, -0.728477, 1.570796, 2.045285],accel_mss,speed_ms,0,blend_radius_m)
  movel([0.473651, -1.512599, -2.471247, -0.728543, 1.570796, 2.044447],accel_mss,speed_ms,0,blend_radius_m)
  movel([0.473950, -1.512766, -2.471095, -0.728527, 1.570796, 2.044746],accel_mss,speed_ms,0,blend_radius_m)
  movel([0.474432, -1.512811, -2.471055, -0.728523, 1.570796, 2.045228],accel_mss,speed_ms,0,blend_radius_m)
  movel([0.475729, -1.512633, -2.471216, -0.728540, 1.570796, 2.046525],accel_mss,speed_ms,0,blend_radius_m)
  movel([0.477102, -1.512257, -2.471557, -0.728575, 1.570796, 2.047899],accel_mss,speed_ms,0,blend_radius_m)
  movel([0.478108, -1.511875, -2.471903, -0.728611, 1.570796, 2.048905],accel_mss,speed_ms,0,blend_radius_m)
  movel([0.478780, -1.511488, -2.472253, -0.728648, 1.570796, 2.049577],accel_mss,speed_ms,0,blend_radius_m)
  movel([0.479133, -1.511140, -2.472568, -0.728681, 1.570796, 2.049929],accel_mss,speed_ms,0,blend_radius_m)
  movel([0.479218, -1.510826, -2.472851, -0.728712, 1.570796, 2.050014],accel_mss,speed_ms,0,blend_radius_m)
  movel([0.479090, -1.510544, -2.473106, -0.728739, 1.570796, 2.049886],accel_mss,speed_ms,0,blend_radius_m)
  movel([0.478414, -1.510068, -2.473536, -0.728785, 1.570796, 2.049210],accel_mss,speed_ms,0,blend_radius_m)
  movel([0.477542, -1.509693, -2.473874, -0.728822, 1.570796, 2.048338],accel_mss,speed_ms,0,blend_radius_m)
  movel([0.475558, -1.508835, -2.474647, -0.728907, 1.570796, 2.046354],accel_mss,speed_ms,0,blend_radius_m)
  movel([0.473690, -1.507767, -2.475608, -0.729014, 1.570796, 2.044487],accel_mss,speed_ms,0,blend_radius_m)
  movel([0.472881, -1.507120, -2.476189, -0.729080, 1.570796, 2.043678],accel_mss,speed_ms,0,blend_radius_m)
  movel([0.472200, -1.506379, -2.476853, -0.729157, 1.570796, 2.042997],accel_mss,speed_ms,0,blend_radius_m)
  movel([0.471682, -1.505529, -2.477615, -0.729245, 1.570796, 2.042478],accel_mss,speed_ms,0,blend_radius_m)
  movel([0.471359, -1.504557, -2.478484, -0.729348, 1.570796, 2.042155],accel_mss,speed_ms,0,blend_radius_m)
  movel([0.472548, -1.505063, -2.478031, -0.729294, 1.570796, 2.043345],accel_mss,speed_ms,0,blend_radius_m)
  movel([0.473290, -1.505166, -2.477940, -0.729283, 1.570796, 2.044086],accel_mss,speed_ms,0,blend_radius_m)
  movel([0.473666, -1.505119, -2.477981, -0.729288, 1.570796, 2.044462],accel_mss,speed_ms,0,blend_radius_m)
  movel([0.474036, -1.504983, -2.478103, -0.729303, 1.570796, 2.044833],accel_mss,speed_ms,0,blend_radius_m)
  movel([0.474250, -1.504808, -2.478260, -0.729321, 1.570796, 2.045046],accel_mss,speed_ms,0,blend_radius_m)
  movel([0.474359, -1.504562, -2.478480, -0.729347, 1.570796, 2.045156],accel_mss,speed_ms,0,blend_radius_m)
  movel([0.474320, -1.503904, -2.479067, -0.729418, 1.570796, 2.045117],accel_mss,speed_ms,0,blend_radius_m)
  movel([0.474008, -1.503088, -2.479795, -0.729506, 1.570796, 2.044804],accel_mss,speed_ms,0,blend_radius_m)
  movel([0.473517, -1.502193, -2.480592, -0.729604, 1.570796, 2.044314],accel_mss,speed_ms,0,blend_radius_m)
  movel([0.471613, -1.499414, -2.483059, -0.729917, 1.570796, 2.042409],accel_mss,speed_ms,0,blend_radius_m)
  movel([0.471030, -1.498202, -2.484130, -0.730057, 1.570796, 2.041827],accel_mss,speed_ms,0,blend_radius_m)
  movel([0.470618, -1.496895, -2.485283, -0.730211, 1.570796, 2.041414],accel_mss,speed_ms,0,blend_radius_m)
  movel([0.470446, -1.495493, -2.486518, -0.730379, 1.570796, 2.041242],accel_mss,speed_ms,0,blend_radius_m)
  movel([0.470580, -1.493993, -2.487834, -0.730562, 1.570796, 2.041377],accel_mss,speed_ms,0,blend_radius_m)
  movel([0.471074, -1.495188, -2.486785, -0.730416, 1.570796, 2.041871],accel_mss,speed_ms,0,blend_radius_m)
  movel([0.471484, -1.495742, -2.486298, -0.730349, 1.570796, 2.042280],accel_mss,speed_ms,0,blend_radius_m)
  movel([0.472012, -1.496033, -2.486042, -0.730314, 1.570796, 2.042808],accel_mss,speed_ms,0,blend_radius_m)
  movel([0.472673, -1.496012, -2.486061, -0.730316, 1.570796, 2.043469],accel_mss,speed_ms,0,blend_radius_m)
  movel([0.473211, -1.495731, -2.486308, -0.730350, 1.570796, 2.044007],accel_mss,speed_ms,0,blend_radius_m)
  movel([0.473577, -1.495256, -2.486726, -0.730407, 1.570796, 2.044373],accel_mss,speed_ms,0,blend_radius_m)
  movel([0.473727, -1.494646, -2.487261, -0.730482, 1.570796, 2.044523],accel_mss,speed_ms,0,blend_radius_m)
  movel([0.473997, -1.491440, -2.490067, -0.730882, 1.570796, 2.044794],accel_mss,speed_ms,0,blend_radius_m)
  movel([0.474620, -1.488224, -2.492866, -0.731299, 1.570796, 2.045417],accel_mss,speed_ms,0,blend_radius_m)
  movel([0.475100, -1.486590, -2.494281, -0.731518, 1.570796, 2.045897],accel_mss,speed_ms,0,blend_radius_m)
  movel([0.475711, -1.484927, -2.495718, -0.731745, 1.570796, 2.046507],accel_mss,speed_ms,0,blend_radius_m)
  movel([0.476467, -1.483225, -2.497183, -0.731981, 1.570796, 2.047263],accel_mss,speed_ms,0,blend_radius_m)
  movel([0.477383, -1.481477, -2.498684, -0.732229, 1.570796, 2.048179],accel_mss,speed_ms,0,blend_radius_m)
  speed_ms = 0.005
  movel([0.477383, -1.473438, -2.495122, -0.743828, 1.570796, 2.048179],accel_mss,speed_ms,0,blend_radius_m)
  speed_ms = 0.040
  movel([0.466032, -1.452408, -2.512575, -0.747407, 1.570796, 2.036828],accel_mss,speed_ms,0,blend_radius_m)
  speed_ms = 0.005
  movel([0.466032, -1.460613, -2.516221, -0.735555, 1.570796, 2.036828],accel_mss,speed_ms,0,blend_radius_m)
  speed_ms = 0.025
  movel([0.468902, -1.458797, -2.517715, -0.735877, 1.570796, 2.039698],accel_mss,speed_ms,0,blend_radius_m)
  movel([0.471734, -1.456911, -2.519262, -0.736216, 1.570796, 2.042530],accel_mss,speed_ms,0,blend_radius_m)
  movel([0.477317, -1.452938, -2.522502, -0.736949, 1.570796, 2.048114],accel_mss,speed_ms,0,blend_radius_m)
  movel([0.482782, -1.448709, -2.525923, -0.737756, 1.570796, 2.053579],accel_mss,speed_ms,0,blend_radius_m)
  movel([0.488116, -1.444241, -2.529509, -0.738639, 1.570796, 2.058913],accel_mss,speed_ms,0,blend_radius_m)
  movel([0.493309, -1.439545, -2.533244, -0.739600, 1.570796, 2.064105],accel_mss,speed_ms,0,blend_radius_m)
  movel([0.498346, -1.434638, -2.537111, -0.740640, 1.570796, 2.069143],accel_mss,speed_ms,0,blend_radius_m)
  movel([0.503214, -1.429536, -2.541092, -0.741760, 1.570796, 2.074011],accel_mss,speed_ms,0,blend_radius_m)
  movel([0.507901, -1.424253, -2.545174, -0.742962, 1.570796, 2.078698],accel_mss,speed_ms,0,blend_radius_m)
  movel([0.512387, -1.418809, -2.549336, -0.744244, 1.570796, 2.083184],accel_mss,speed_ms,0,blend_radius_m)
  movel([0.516658, -1.413219, -2.553563, -0.745607, 1.570796, 2.087454],accel_mss,speed_ms,0,blend_radius_m)
  movel([0.520693, -1.407501, -2.557838, -0.747050, 1.570796, 2.091490],accel_mss,speed_ms,0,blend_radius_m)
  movel([0.524474, -1.401675, -2.562144, -0.748570, 1.570796, 2.095271],accel_mss,speed_ms,0,blend_radius_m)
  movel([0.527986, -1.395759, -2.566466, -0.750164, 1.570796, 2.098783],accel_mss,speed_ms,0,blend_radius_m)
  movel([0.531202, -1.389774, -2.570785, -0.751829, 1.570796, 2.101998],accel_mss,speed_ms,0,blend_radius_m)
  movel([0.534102, -1.383745, -2.575084, -0.753560, 1.570796, 2.104898],accel_mss,speed_ms,0,blend_radius_m)
  movel([0.537945, -1.374648, -2.581470, -0.756271, 1.570796, 2.108741],accel_mss,speed_ms,0,blend_radius_m)
  movel([0.538771, -1.373143, -2.582516, -0.756731, 1.570796, 2.109567],accel_mss,speed_ms,0,blend_radius_m)
  movel([0.539817, -1.371681, -2.583528, -0.757181, 1.570796, 2.110613],accel_mss,speed_ms,0,blend_radius_m)
  movel([0.541538, -1.369792, -2.584831, -0.757767, 1.570796, 2.112334],accel_mss,speed_ms,0,blend_radius_m)
  movel([0.543091, -1.368476, -2.585735, -0.758178, 1.570796, 2.113887],accel_mss,speed_ms,0,blend_radius_m)
  movel([0.543804, -1.368020, -2.586049, -0.758321, 1.570796, 2.114601],accel_mss,speed_ms,0,blend_radius_m)
  movel([0.545113, -1.367469, -2.586426, -0.758494, 1.570796, 2.115909],accel_mss,speed_ms,0,blend_radius_m)
  movel([0.545705, -1.367366, -2.586497, -0.758526, 1.570796, 2.116501],accel_mss,speed_ms,0,blend_radius_m)
  movel([0.546777, -1.367466, -2.586428, -0.758495, 1.570796, 2.117574],accel_mss,speed_ms,0,blend_radius_m)
  movel([0.547701, -1.367929, -2.586111, -0.758349, 1.570796, 2.118497],accel_mss,speed_ms,0,blend_radius_m)
  movel([0.548483, -1.368700, -2.585581, -0.758107, 1.570796, 2.119280],accel_mss,speed_ms,0,blend_radius_m)
  movel([0.549132, -1.369728, -2.584875, -0.757786, 1.570796, 2.119928],accel_mss,speed_ms,0,blend_radius_m)
  movel([0.549655, -1.370952, -2.584031, -0.757406, 1.570796, 2.120452],accel_mss,speed_ms,0,blend_radius_m)
  movel([0.550060, -1.372322, -2.583084, -0.756983, 1.570796, 2.120856],accel_mss,speed_ms,0,blend_radius_m)
  movel([0.550551, -1.375266, -2.581040, -0.756083, 1.570796, 2.121347],accel_mss,speed_ms,0,blend_radius_m)
  movel([0.550668, -1.378132, -2.579039, -0.755219, 1.570796, 2.121464],accel_mss,speed_ms,0,blend_radius_m)
  movel([0.550484, -1.380487, -2.577385, -0.754517, 1.570796, 2.121281],accel_mss,speed_ms,0,blend_radius_m)
  movel([0.549919, -1.383302, -2.575398, -0.753689, 1.570796, 2.120715],accel_mss,speed_ms,0,blend_radius_m)
  movel([0.549155, -1.386148, -2.573377, -0.752864, 1.570796, 2.119951],accel_mss,speed_ms,0,blend_radius_m)
  movel([0.547245, -1.391873, -2.569277, -0.751240, 1.570796, 2.118042],accel_mss,speed_ms,0,blend_radius_m)
  movel([0.545162, -1.397558, -2.565157, -0.749674, 1.570796, 2.115959],accel_mss,speed_ms,0,blend_radius_m)
  movel([0.543302, -1.403099, -2.561096, -0.748194, 1.570796, 2.114098],accel_mss,speed_ms,0,blend_radius_m)
  movel([0.541964, -1.407989, -2.557475, -0.746925, 1.570796, 2.112760],accel_mss,speed_ms,0,blend_radius_m)
  movel([0.541538, -1.410366, -2.555702, -0.746321, 1.570796, 2.112334],accel_mss,speed_ms,0,blend_radius_m)
  movel([0.541409, -1.412652, -2.553988, -0.745748, 1.570796, 2.112205],accel_mss,speed_ms,0,blend_radius_m)
  movel([0.541530, -1.413653, -2.553236, -0.745500, 1.570796, 2.112327],accel_mss,speed_ms,0,blend_radius_m)
  movel([0.541712, -1.414085, -2.552911, -0.745393, 1.570796, 2.112508],accel_mss,speed_ms,0,blend_radius_m)
  movel([0.542014, -1.414430, -2.552651, -0.745308, 1.570796, 2.112811],accel_mss,speed_ms,0,blend_radius_m)
  movel([0.542579, -1.414692, -2.552453, -0.745244, 1.570796, 2.113375],accel_mss,speed_ms,0,blend_radius_m)
  movel([0.543278, -1.414768, -2.552396, -0.745225, 1.570796, 2.114074],accel_mss,speed_ms,0,blend_radius_m)
  movel([0.544866, -1.414552, -2.552559, -0.745278, 1.570796, 2.115662],accel_mss,speed_ms,0,blend_radius_m)
  movel([0.546735, -1.414053, -2.552935, -0.745401, 1.570796, 2.117531],accel_mss,speed_ms,0,blend_radius_m)
  movel([0.548597, -1.413416, -2.553414, -0.745558, 1.570796, 2.119394],accel_mss,speed_ms,0,blend_radius_m)
  movel([0.552310, -1.411832, -2.554605, -0.745953, 1.570796, 2.123106],accel_mss,speed_ms,0,blend_radius_m)
  movel([0.559726, -1.408243, -2.557286, -0.746860, 1.570796, 2.130523],accel_mss,speed_ms,0,blend_radius_m)
  movel([0.563228, -1.406710, -2.558426, -0.747253, 1.570796, 2.134025],accel_mss,speed_ms,0,blend_radius_m)
  movel([0.565185, -1.405992, -2.558959, -0.747439, 1.570796, 2.135981],accel_mss,speed_ms,0,blend_radius_m)
  movel([0.567041, -1.405492, -2.559329, -0.747568, 1.570796, 2.137837],accel_mss,speed_ms,0,blend_radius_m)
  movel([0.567877, -1.405366, -2.559422, -0.747601, 1.570796, 2.138673],accel_mss,speed_ms,0,blend_radius_m)
  movel([0.568623, -1.405347, -2.559436, -0.747606, 1.570796, 2.139419],accel_mss,speed_ms,0,blend_radius_m)
  movel([0.569256, -1.405450, -2.559360, -0.747579, 1.570796, 2.140052],accel_mss,speed_ms,0,blend_radius_m)
  movel([0.569753, -1.405695, -2.559178, -0.747516, 1.570796, 2.140549],accel_mss,speed_ms,0,blend_radius_m)
  movel([0.570094, -1.406095, -2.558882, -0.747412, 1.570796, 2.140890],accel_mss,speed_ms,0,blend_radius_m)
  movel([0.570258, -1.406668, -2.558457, -0.747264, 1.570796, 2.141054],accel_mss,speed_ms,0,blend_radius_m)
  movel([0.570222, -1.407432, -2.557890, -0.747068, 1.570796, 2.141018],accel_mss,speed_ms,0,blend_radius_m)
  movel([0.569963, -1.408401, -2.557168, -0.746820, 1.570796, 2.140760],accel_mss,speed_ms,0,blend_radius_m)
  movel([0.569286, -1.410124, -2.555883, -0.746382, 1.570796, 2.140083],accel_mss,speed_ms,0,blend_radius_m)
  movel([0.568475, -1.411800, -2.554629, -0.745961, 1.570796, 2.139271],accel_mss,speed_ms,0,blend_radius_m)
  movel([0.567540, -1.413425, -2.553408, -0.745556, 1.570796, 2.138336],accel_mss,speed_ms,0,blend_radius_m)
  movel([0.566489, -1.415003, -2.552219, -0.745167, 1.570796, 2.137285],accel_mss,speed_ms,0,blend_radius_m)
  movel([0.565332, -1.416528, -2.551066, -0.744795, 1.570796, 2.136128],accel_mss,speed_ms,0,blend_radius_m)
  movel([0.564077, -1.418002, -2.549949, -0.744438, 1.570796, 2.134873],accel_mss,speed_ms,0,blend_radius_m)
  movel([0.562731, -1.419423, -2.548869, -0.744097, 1.570796, 2.133528],accel_mss,speed_ms,0,blend_radius_m)
  movel([0.561305, -1.420792, -2.547825, -0.743772, 1.570796, 2.132101],accel_mss,speed_ms,0,blend_radius_m)
  movel([0.558245, -1.423366, -2.545855, -0.743168, 1.570796, 2.129041],accel_mss,speed_ms,0,blend_radius_m)
  movel([0.554959, -1.425720, -2.544045, -0.742624, 1.570796, 2.125756],accel_mss,speed_ms,0,blend_radius_m)
  movel([0.551512, -1.427846, -2.542403, -0.742140, 1.570796, 2.122308],accel_mss,speed_ms,0,blend_radius_m)
  movel([0.547970, -1.429739, -2.540935, -0.741715, 1.570796, 2.118766],accel_mss,speed_ms,0,blend_radius_m)
  movel([0.539979, -1.433664, -2.537874, -0.740851, 1.570796, 2.110775],accel_mss,speed_ms,0,blend_radius_m)
  movel([0.535909, -1.435398, -2.536514, -0.740477, 1.570796, 2.106705],accel_mss,speed_ms,0,blend_radius_m)
  movel([0.533914, -1.436111, -2.535954, -0.740324, 1.570796, 2.104710],accel_mss,speed_ms,0,blend_radius_m)
  movel([0.531965, -1.436684, -2.535503, -0.740202, 1.570796, 2.102762],accel_mss,speed_ms,0,blend_radius_m)
  movel([0.530749, -1.436952, -2.535292, -0.740145, 1.570796, 2.101545],accel_mss,speed_ms,0,blend_radius_m)
  movel([0.529585, -1.437111, -2.535167, -0.740111, 1.570796, 2.100382],accel_mss,speed_ms,0,blend_radius_m)
  movel([0.528488, -1.437147, -2.535138, -0.740104, 1.570796, 2.099284],accel_mss,speed_ms,0,blend_radius_m)
  movel([0.527472, -1.437051, -2.535214, -0.740124, 1.570796, 2.098268],accel_mss,speed_ms,0,blend_radius_m)
  movel([0.526552, -1.436813, -2.535401, -0.740174, 1.570796, 2.097349],accel_mss,speed_ms,0,blend_radius_m)
  movel([0.525742, -1.436422, -2.535709, -0.740258, 1.570796, 2.096539],accel_mss,speed_ms,0,blend_radius_m)
  movel([0.525060, -1.435863, -2.536149, -0.740377, 1.570796, 2.095857],accel_mss,speed_ms,0,blend_radius_m)
  movel([0.524520, -1.435125, -2.536729, -0.740535, 1.570796, 2.095316],accel_mss,speed_ms,0,blend_radius_m)
  movel([0.524155, -1.434223, -2.537437, -0.740730, 1.570796, 2.094952],accel_mss,speed_ms,0,blend_radius_m)
  movel([0.523975, -1.433243, -2.538203, -0.740942, 1.570796, 2.094772],accel_mss,speed_ms,0,blend_radius_m)
  movel([0.523875, -1.429029, -2.541486, -0.741874, 1.570796, 2.094671],accel_mss,speed_ms,0,blend_radius_m)
  movel([0.523695, -1.428021, -2.542268, -0.742101, 1.570796, 2.094491],accel_mss,speed_ms,0,blend_radius_m)
  movel([0.523325, -1.427082, -2.542994, -0.742313, 1.570796, 2.094122],accel_mss,speed_ms,0,blend_radius_m)
  movel([0.523071, -1.426813, -2.543202, -0.742374, 1.570796, 2.093867],accel_mss,speed_ms,0,blend_radius_m)
  movel([0.522822, -1.426930, -2.543111, -0.742348, 1.570796, 2.093618],accel_mss,speed_ms,0,blend_radius_m)
  movel([0.522355, -1.427345, -2.542790, -0.742254, 1.570796, 2.093151],accel_mss,speed_ms,0,blend_radius_m)
  movel([0.520874, -1.428916, -2.541574, -0.741899, 1.570796, 2.091670],accel_mss,speed_ms,0,blend_radius_m)
  movel([0.516616, -1.433877, -2.537707, -0.740805, 1.570796, 2.087413],accel_mss,speed_ms,0,blend_radius_m)
  movel([0.509629, -1.442253, -2.531094, -0.739042, 1.570796, 2.080425],accel_mss,speed_ms,0,blend_radius_m)
  movel([0.505584, -1.446410, -2.527772, -0.738207, 1.570796, 2.076380],accel_mss,speed_ms,0,blend_radius_m)
  movel([0.501403, -1.450431, -2.524534, -0.737424, 1.570796, 2.072199],accel_mss,speed_ms,0,blend_radius_m)
  movel([0.497105, -1.454321, -2.521377, -0.736691, 1.570796, 2.067901],accel_mss,speed_ms,0,blend_radius_m)
  movel([0.492719, -1.458086, -2.518299, -0.736004, 1.570796, 2.063515],accel_mss,speed_ms,0,blend_radius_m)
  movel([0.487033, -1.462788, -2.514425, -0.735177, 1.570796, 2.057830],accel_mss,speed_ms,0,blend_radius_m)
  movel([0.481276, -1.467394, -2.510596, -0.734399, 1.570796, 2.052072],accel_mss,speed_ms,0,blend_radius_m)
  movel([0.475444, -1.471860, -2.506851, -0.733677, 1.570796, 2.046241],accel_mss,speed_ms,0,blend_radius_m)
  movel([0.469530, -1.476139, -2.503235, -0.733015, 1.570796, 2.040326],accel_mss,speed_ms,0,blend_radius_m)
  movel([0.463529, -1.480182, -2.499792, -0.732415, 1.570796, 2.034326],accel_mss,speed_ms,0,blend_radius_m)
  movel([0.460496, -1.482104, -2.498146, -0.732139, 1.570796, 2.031292],accel_mss,speed_ms,0,blend_radius_m)
  movel([0.457435, -1.483950, -2.496559, -0.731880, 1.570796, 2.028231],accel_mss,speed_ms,0,blend_radius_m)
  movel([0.454348, -1.485717, -2.495035, -0.731636, 1.570796, 2.025144],accel_mss,speed_ms,0,blend_radius_m)
  movel([0.451235, -1.487398, -2.493582, -0.731409, 1.570796, 2.022032],accel_mss,speed_ms,0,blend_radius_m)
  movel([0.448093, -1.488991, -2.492200, -0.731198, 1.570796, 2.018889],accel_mss,speed_ms,0,blend_radius_m)
  movel([0.444920, -1.490485, -2.490900, -0.731004, 1.570796, 2.015717],accel_mss,speed_ms,0,blend_radius_m)
  movel([0.441121, -1.492138, -2.489458, -0.730793, 1.570796, 2.011917],accel_mss,speed_ms,0,blend_radius_m)
  movel([0.439214, -1.492856, -2.488830, -0.730703, 1.570796, 2.010010],accel_mss,speed_ms,0,blend_radius_m)
  movel([0.435953, -1.493815, -2.487990, -0.730584, 1.570796, 2.006750],accel_mss,speed_ms,0,blend_radius_m)
  movel([0.434355, -1.494140, -2.487706, -0.730544, 1.570796, 2.005151],accel_mss,speed_ms,0,blend_radius_m)
  movel([0.432892, -1.494199, -2.487654, -0.730536, 1.570796, 2.003689],accel_mss,speed_ms,0,blend_radius_m)
  movel([0.432332, -1.494057, -2.487778, -0.730554, 1.570796, 2.003129],accel_mss,speed_ms,0,blend_radius_m)
  movel([0.431947, -1.493762, -2.488037, -0.730590, 1.570796, 2.002743],accel_mss,speed_ms,0,blend_radius_m)
  movel([0.433050, -1.492467, -2.489170, -0.730752, 1.570796, 2.003846],accel_mss,speed_ms,0,blend_radius_m)
  movel([0.433977, -1.491111, -2.490354, -0.730924, 1.570796, 2.004774],accel_mss,speed_ms,0,blend_radius_m)
  movel([0.434304, -1.490444, -2.490936, -0.731009, 1.570796, 2.005100],accel_mss,speed_ms,0,blend_radius_m)
  movel([0.434501, -1.489802, -2.491495, -0.731092, 1.570796, 2.005297],accel_mss,speed_ms,0,blend_radius_m)
  movel([0.434541, -1.489197, -2.492021, -0.731171, 1.570796, 2.005338],accel_mss,speed_ms,0,blend_radius_m)
  movel([0.434390, -1.488645, -2.492501, -0.731244, 1.570796, 2.005186],accel_mss,speed_ms,0,blend_radius_m)
  movel([0.433605, -1.487527, -2.493470, -0.731392, 1.570796, 2.004401],accel_mss,speed_ms,0,blend_radius_m)
  movel([0.433481, -1.487048, -2.493885, -0.731456, 1.570796, 2.004278],accel_mss,speed_ms,0,blend_radius_m)
  movel([0.433504, -1.486523, -2.494339, -0.731527, 1.570796, 2.004300],accel_mss,speed_ms,0,blend_radius_m)
  movel([0.433910, -1.485389, -2.495318, -0.731681, 1.570796, 2.004706],accel_mss,speed_ms,0,blend_radius_m)
  movel([0.434649, -1.484208, -2.496337, -0.731844, 1.570796, 2.005445],accel_mss,speed_ms,0,blend_radius_m)
  movel([0.435548, -1.483069, -2.497317, -0.732003, 1.570796, 2.006344],accel_mss,speed_ms,0,blend_radius_m)
  movel([0.438447, -1.479730, -2.500178, -0.732481, 1.570796, 2.009243],accel_mss,speed_ms,0,blend_radius_m)
  movel([0.441555, -1.476440, -2.502980, -0.732969, 1.570796, 2.012351],accel_mss,speed_ms,0,blend_radius_m)
  movel([0.443204, -1.474853, -2.504325, -0.733211, 1.570796, 2.014000],accel_mss,speed_ms,0,blend_radius_m)
  movel([0.444924, -1.473320, -2.505621, -0.733448, 1.570796, 2.015721],accel_mss,speed_ms,0,blend_radius_m)
  movel([0.446722, -1.471861, -2.506851, -0.733677, 1.570796, 2.017518],accel_mss,speed_ms,0,blend_radius_m)
  movel([0.448605, -1.470491, -2.508003, -0.733895, 1.570796, 2.019402],accel_mss,speed_ms,0,blend_radius_m)
  movel([0.450533, -1.469313, -2.508991, -0.734085, 1.570796, 2.021329],accel_mss,speed_ms,0,blend_radius_m)
  movel([0.456408, -1.466369, -2.511451, -0.734569, 1.570796, 2.027205],accel_mss,speed_ms,0,blend_radius_m)
  movel([0.461233, -1.463560, -2.513785, -0.735044, 1.570796, 2.032030],accel_mss,speed_ms,0,blend_radius_m)
  movel([0.466032, -1.460613, -2.516221, -0.735555, 1.570796, 2.036828],accel_mss,speed_ms,0,blend_radius_m)
  movel([0.468181, -1.459252, -2.517341, -0.735796, 1.570796, 2.038977],accel_mss,speed_ms,0,blend_radius_m)
  speed_ms = 0.005
  movel([0.468181, -1.451036, -2.513689, -0.747664, 1.570796, 2.038977],accel_mss,speed_ms,0,blend_radius_m)
  speed_ms = 0.040
  movel([0.426259, -1.473575, -2.495006, -0.743807, 1.570796, 1.997056],accel_mss,speed_ms,0,blend_radius_m)
  speed_ms = 0.005
  movel([0.426259, -1.481613, -2.498567, -0.732209, 1.570796, 1.997056],accel_mss,speed_ms,0,blend_radius_m)
  speed_ms = 0.025
  movel([0.426785, -1.485296, -2.495399, -0.731694, 1.570796, 1.997582],accel_mss,speed_ms,0,blend_radius_m)
  movel([0.426943, -1.487302, -2.493665, -0.731422, 1.570796, 1.997739],accel_mss,speed_ms,0,blend_radius_m)
  movel([0.426956, -1.489374, -2.491867, -0.731148, 1.570796, 1.997753],accel_mss,speed_ms,0,blend_radius_m)
  movel([0.426780, -1.491475, -2.490037, -0.730877, 1.570796, 1.997576],accel_mss,speed_ms,0,blend_radius_m)
  movel([0.426361, -1.493570, -2.488205, -0.730614, 1.570796, 1.997157],accel_mss,speed_ms,0,blend_radius_m)
  movel([0.425648, -1.495628, -2.486399, -0.730362, 1.570796, 1.996444],accel_mss,speed_ms,0,blend_radius_m)
  movel([0.425164, -1.496634, -2.485513, -0.730242, 1.570796, 1.995961],accel_mss,speed_ms,0,blend_radius_m)
  movel([0.424590, -1.497615, -2.484648, -0.730126, 1.570796, 1.995386],accel_mss,speed_ms,0,blend_radius_m)
  movel([0.424302, -1.496994, -2.485196, -0.730199, 1.570796, 1.995098],accel_mss,speed_ms,0,blend_radius_m)
  movel([0.424245, -1.496354, -2.485760, -0.730275, 1.570796, 1.995041],accel_mss,speed_ms,0,blend_radius_m)
  movel([0.424185, -1.494900, -2.487039, -0.730451, 1.570796, 1.994982],accel_mss,speed_ms,0,blend_radius_m)
  movel([0.423788, -1.493467, -2.488295, -0.730627, 1.570796, 1.994585],accel_mss,speed_ms,0,blend_radius_m)
  movel([0.423223, -1.492114, -2.489479, -0.730796, 1.570796, 1.994019],accel_mss,speed_ms,0,blend_radius_m)
  movel([0.422503, -1.490843, -2.490588, -0.730958, 1.570796, 1.993300],accel_mss,speed_ms,0,blend_radius_m)
  movel([0.421640, -1.489659, -2.491619, -0.731111, 1.570796, 1.992436],accel_mss,speed_ms,0,blend_radius_m)
  movel([0.420645, -1.488568, -2.492567, -0.731254, 1.570796, 1.991442],accel_mss,speed_ms,0,blend_radius_m)
  movel([0.419531, -1.487577, -2.493427, -0.731385, 1.570796, 1.990327],accel_mss,speed_ms,0,blend_radius_m)
  movel([0.418306, -1.486690, -2.494195, -0.731504, 1.570796, 1.989103],accel_mss,speed_ms,0,blend_radius_m)
  movel([0.416988, -1.485911, -2.494868, -0.731610, 1.570796, 1.987784],accel_mss,speed_ms,0,blend_radius_m)
  movel([0.416041, -1.485484, -2.495237, -0.731668, 1.570796, 1.986838],accel_mss,speed_ms,0,blend_radius_m)
  movel([0.415222, -1.485270, -2.495421, -0.731697, 1.570796, 1.986019],accel_mss,speed_ms,0,blend_radius_m)
  movel([0.414524, -1.485248, -2.495440, -0.731700, 1.570796, 1.985320],accel_mss,speed_ms,0,blend_radius_m)
  movel([0.413938, -1.485397, -2.495312, -0.731680, 1.570796, 1.984734],accel_mss,speed_ms,0,blend_radius_m)
  movel([0.413451, -1.485701, -2.495049, -0.731638, 1.570796, 1.984247],accel_mss,speed_ms,0,blend_radius_m)
  movel([0.413056, -1.486139, -2.494671, -0.731579, 1.570796, 1.983852],accel_mss,speed_ms,0,blend_radius_m)
  movel([0.412740, -1.486691, -2.494194, -0.731504, 1.570796, 1.983536],accel_mss,speed_ms,0,blend_radius_m)
  movel([0.412496, -1.487338, -2.493634, -0.731417, 1.570796, 1.983292],accel_mss,speed_ms,0,blend_radius_m)
  movel([0.412176, -1.488839, -2.492331, -0.731218, 1.570796, 1.982973],accel_mss,speed_ms,0,blend_radius_m)
  movel([0.411827, -1.493652, -2.488133, -0.730604, 1.570796, 1.982623],accel_mss,speed_ms,0,blend_radius_m)
  movel([0.411194, -1.492016, -2.489564, -0.730809, 1.570796, 1.981990],accel_mss,speed_ms,0,blend_radius_m)
  movel([0.410024, -1.488695, -2.492457, -0.731237, 1.570796, 1.980820],accel_mss,speed_ms,0,blend_radius_m)
  movel([0.409157, -1.487197, -2.493756, -0.731436, 1.570796, 1.979953],accel_mss,speed_ms,0,blend_radius_m)
  movel([0.407933, -1.485717, -2.495036, -0.731636, 1.570796, 1.978730],accel_mss,speed_ms,0,blend_radius_m)
  movel([0.406592, -1.484312, -2.496248, -0.731830, 1.570796, 1.977388],accel_mss,speed_ms,0,blend_radius_m)
  movel([0.403823, -1.481556, -2.498615, -0.732217, 1.570796, 1.974619],accel_mss,speed_ms,0,blend_radius_m)
  movel([0.402529, -1.480121, -2.499844, -0.732424, 1.570796, 1.973326],accel_mss,speed_ms,0,blend_radius_m)
  movel([0.401388, -1.478591, -2.501149, -0.732648, 1.570796, 1.972184],accel_mss,speed_ms,0,blend_radius_m)
  movel([0.400466, -1.476926, -2.502567, -0.732896, 1.570796, 1.971262],accel_mss,speed_ms,0,blend_radius_m)
  movel([0.399832, -1.475077, -2.504136, -0.733177, 1.570796, 1.970629],accel_mss,speed_ms,0,blend_radius_m)
  movel([0.399145, -1.479131, -2.500689, -0.732569, 1.570796, 1.969941],accel_mss,speed_ms,0,blend_radius_m)
  movel([0.398904, -1.481187, -2.498932, -0.732270, 1.570796, 1.969701],accel_mss,speed_ms,0,blend_radius_m)
  movel([0.398906, -1.483032, -2.497348, -0.732008, 1.570796, 1.969703],accel_mss,speed_ms,0,blend_radius_m)
  movel([0.398200, -1.481266, -2.498864, -0.732259, 1.570796, 1.968996],accel_mss,speed_ms,0,blend_radius_m)
  movel([0.397271, -1.479624, -2.500269, -0.732497, 1.570796, 1.968068],accel_mss,speed_ms,0,blend_radius_m)
  movel([0.395194, -1.476458, -2.502964, -0.732967, 1.570796, 1.965991],accel_mss,speed_ms,0,blend_radius_m)
  movel([0.394608, -1.475326, -2.503925, -0.733139, 1.570796, 1.965405],accel_mss,speed_ms,0,blend_radius_m)
  movel([0.394185, -1.474140, -2.504928, -0.733321, 1.570796, 1.964981],accel_mss,speed_ms,0,blend_radius_m)
  movel([0.393661, -1.471651, -2.507028, -0.733710, 1.570796, 1.964457],accel_mss,speed_ms,0,blend_radius_m)
  movel([0.393279, -1.469083, -2.509184, -0.734123, 1.570796, 1.964076],accel_mss,speed_ms,0,blend_radius_m)
  movel([0.392690, -1.466536, -2.511311, -0.734542, 1.570796, 1.963486],accel_mss,speed_ms,0,blend_radius_m)
  movel([0.392390, -1.465786, -2.511936, -0.734667, 1.570796, 1.963186],accel_mss,speed_ms,0,blend_radius_m)
  movel([0.391952, -1.465122, -2.512488, -0.734778, 1.570796, 1.962748],accel_mss,speed_ms,0,blend_radius_m)
  movel([0.391326, -1.464651, -2.512880, -0.734858, 1.570796, 1.962122],accel_mss,speed_ms,0,blend_radius_m)
  movel([0.390931, -1.464520, -2.512989, -0.734880, 1.570796, 1.961727],accel_mss,speed_ms,0,blend_radius_m)
  movel([0.390469, -1.464478, -2.513023, -0.734887, 1.570796, 1.961266],accel_mss,speed_ms,0,blend_radius_m)
  movel([0.389918, -1.464541, -2.512972, -0.734877, 1.570796, 1.960714],accel_mss,speed_ms,0,blend_radius_m)
  movel([0.389364, -1.464708, -2.512833, -0.734849, 1.570796, 1.960160],accel_mss,speed_ms,0,blend_radius_m)
  movel([0.388261, -1.465288, -2.512351, -0.734751, 1.570796, 1.959057],accel_mss,speed_ms,0,blend_radius_m)
  movel([0.387204, -1.466087, -2.511686, -0.734616, 1.570796, 1.958001],accel_mss,speed_ms,0,blend_radius_m)
  movel([0.386238, -1.466975, -2.510946, -0.734469, 1.570796, 1.957034],accel_mss,speed_ms,0,blend_radius_m)
  movel([0.386761, -1.465043, -2.512554, -0.734792, 1.570796, 1.957557],accel_mss,speed_ms,0,blend_radius_m)
  movel([0.387114, -1.463166, -2.514112, -0.735111, 1.570796, 1.957911],accel_mss,speed_ms,0,blend_radius_m)
  movel([0.387493, -1.459519, -2.517122, -0.735748, 1.570796, 1.958289],accel_mss,speed_ms,0,blend_radius_m)
  movel([0.387757, -1.455899, -2.520090, -0.736401, 1.570796, 1.958553],accel_mss,speed_ms,0,blend_radius_m)
  movel([0.388297, -1.452167, -2.523127, -0.737094, 1.570796, 1.959094],accel_mss,speed_ms,0,blend_radius_m)
  movel([0.388714, -1.450679, -2.524333, -0.737377, 1.570796, 1.959510],accel_mss,speed_ms,0,blend_radius_m)
  movel([0.389333, -1.449137, -2.525579, -0.737674, 1.570796, 1.960129],accel_mss,speed_ms,0,blend_radius_m)
  movel([0.390119, -1.447559, -2.526849, -0.737981, 1.570796, 1.960915],accel_mss,speed_ms,0,blend_radius_m)
  movel([0.391033, -1.445967, -2.528127, -0.738295, 1.570796, 1.961829],accel_mss,speed_ms,0,blend_radius_m)
  movel([0.393120, -1.442815, -2.530647, -0.738927, 1.570796, 1.963916],accel_mss,speed_ms,0,blend_radius_m)
  movel([0.395304, -1.439843, -2.533008, -0.739538, 1.570796, 1.966100],accel_mss,speed_ms,0,blend_radius_m)
  speed_ms = 0.005
  movel([0.395304, -1.431474, -2.529275, -0.751640, 1.570796, 1.966100],accel_mss,speed_ms,0,blend_radius_m)
  speed_ms = 0.040
  # Splitting Linear movement in 2 (instruction 806: MoveL 765)
  movel([0.433547, -1.397430, -2.555032, -0.759927, 1.570796, 2.004344],accel_mss,speed_ms,0,blend_radius_m)
  movel([0.474434, -1.362082, -2.579990, -0.770317, 1.570796, 2.045231],accel_mss,speed_ms,0,blend_radius_m)
  speed_ms = 0.005
  movel([0.474434, -1.370965, -2.584022, -0.757402, 1.570796, 2.045231],accel_mss,speed_ms,0,blend_radius_m)
  speed_ms = 0.025
  movel([0.472989, -1.371456, -2.583683, -0.757250, 1.570796, 2.043785],accel_mss,speed_ms,0,blend_radius_m)
  movel([0.472799, -1.371633, -2.583560, -0.757195, 1.570796, 2.043595],accel_mss,speed_ms,0,blend_radius_m)
  movel([0.472675, -1.372000, -2.583307, -0.757082, 1.570796, 2.043471],accel_mss,speed_ms,0,blend_radius_m)
  movel([0.472603, -1.373262, -2.582433, -0.756694, 1.570796, 2.043400],accel_mss,speed_ms,0,blend_radius_m)
  movel([0.473061, -1.377529, -2.579460, -0.755399, 1.570796, 2.043857],accel_mss,speed_ms,0,blend_radius_m)
  movel([0.474120, -1.383440, -2.575300, -0.753649, 1.570796, 2.044916],accel_mss,speed_ms,0,blend_radius_m)
  movel([0.475543, -1.390187, -2.570489, -0.751713, 1.570796, 2.046339],accel_mss,speed_ms,0,blend_radius_m)
  movel([0.478558, -1.403067, -2.561120, -0.748202, 1.570796, 2.049354],accel_mss,speed_ms,0,blend_radius_m)
  movel([0.480397, -1.410133, -2.555876, -0.746380, 1.570796, 2.051193],accel_mss,speed_ms,0,blend_radius_m)
  movel([0.480639, -1.410710, -2.555445, -0.746234, 1.570796, 2.051436],accel_mss,speed_ms,0,blend_radius_m)
  movel([0.481007, -1.411202, -2.555076, -0.746111, 1.570796, 2.051803],accel_mss,speed_ms,0,blend_radius_m)
  movel([0.481528, -1.411486, -2.554864, -0.746039, 1.570796, 2.052324],accel_mss,speed_ms,0,blend_radius_m)
  movel([0.481855, -1.411515, -2.554842, -0.746032, 1.570796, 2.052651],accel_mss,speed_ms,0,blend_radius_m)
  movel([0.482232, -1.411444, -2.554895, -0.746050, 1.570796, 2.053028],accel_mss,speed_ms,0,blend_radius_m)
  movel([0.482920, -1.411095, -2.555156, -0.746137, 1.570796, 2.053716],accel_mss,speed_ms,0,blend_radius_m)
  movel([0.483556, -1.410598, -2.555529, -0.746263, 1.570796, 2.054352],accel_mss,speed_ms,0,blend_radius_m)
  movel([0.486901, -1.407573, -2.557785, -0.747032, 1.570796, 2.057697],accel_mss,speed_ms,0,blend_radius_m)
  movel([0.490066, -1.404379, -2.560152, -0.747858, 1.570796, 2.060862],accel_mss,speed_ms,0,blend_radius_m)
  movel([0.493048, -1.401044, -2.562608, -0.748737, 1.570796, 2.063844],accel_mss,speed_ms,0,blend_radius_m)
  movel([0.495856, -1.397597, -2.565129, -0.749663, 1.570796, 2.066652],accel_mss,speed_ms,0,blend_radius_m)
  movel([0.498491, -1.394061, -2.567697, -0.750631, 1.570796, 2.069287],accel_mss,speed_ms,0,blend_radius_m)
  movel([0.500957, -1.390465, -2.570289, -0.751635, 1.570796, 2.071754],accel_mss,speed_ms,0,blend_radius_m)
  movel([0.503258, -1.386836, -2.572887, -0.752666, 1.570796, 2.074055],accel_mss,speed_ms,0,blend_radius_m)
  movel([0.505395, -1.383207, -2.575465, -0.753717, 1.570796, 2.076191],accel_mss,speed_ms,0,blend_radius_m)
  movel([0.506270, -1.381540, -2.576643, -0.754206, 1.570796, 2.077066],accel_mss,speed_ms,0,blend_radius_m)
  movel([0.506956, -1.379963, -2.577753, -0.754673, 1.570796, 2.077752],accel_mss,speed_ms,0,blend_radius_m)
  movel([0.507455, -1.378474, -2.578799, -0.755116, 1.570796, 2.078251],accel_mss,speed_ms,0,blend_radius_m)
  movel([0.507775, -1.377073, -2.579780, -0.755537, 1.570796, 2.078572],accel_mss,speed_ms,0,blend_radius_m)
  movel([0.507919, -1.375760, -2.580696, -0.755933, 1.570796, 2.078715],accel_mss,speed_ms,0,blend_radius_m)
  movel([0.507889, -1.374537, -2.581547, -0.756305, 1.570796, 2.078686],accel_mss,speed_ms,0,blend_radius_m)
  movel([0.507696, -1.373399, -2.582338, -0.756652, 1.570796, 2.078492],accel_mss,speed_ms,0,blend_radius_m)
  movel([0.507340, -1.372345, -2.583068, -0.756976, 1.570796, 2.078137],accel_mss,speed_ms,0,blend_radius_m)
  movel([0.506829, -1.371378, -2.583737, -0.757274, 1.570796, 2.077625],accel_mss,speed_ms,0,blend_radius_m)
  movel([0.506167, -1.370497, -2.584345, -0.757547, 1.570796, 2.076963],accel_mss,speed_ms,0,blend_radius_m)
  movel([0.505358, -1.369697, -2.584896, -0.757796, 1.570796, 2.076154],accel_mss,speed_ms,0,blend_radius_m)
  movel([0.504410, -1.368982, -2.585388, -0.758019, 1.570796, 2.075207],accel_mss,speed_ms,0,blend_radius_m)
  movel([0.502113, -1.367799, -2.586200, -0.758390, 1.570796, 2.072910],accel_mss,speed_ms,0,blend_radius_m)
  movel([0.499324, -1.366940, -2.586788, -0.758661, 1.570796, 2.070120],accel_mss,speed_ms,0,blend_radius_m)
  movel([0.496587, -1.366526, -2.587072, -0.758791, 1.570796, 2.067383],accel_mss,speed_ms,0,blend_radius_m)
  movel([0.493687, -1.366467, -2.587112, -0.758810, 1.570796, 2.064483],accel_mss,speed_ms,0,blend_radius_m)
  movel([0.490645, -1.366722, -2.586938, -0.758729, 1.570796, 2.061441],accel_mss,speed_ms,0,blend_radius_m)
  movel([0.487496, -1.367238, -2.586584, -0.758567, 1.570796, 2.058292],accel_mss,speed_ms,0,blend_radius_m)
  movel([0.484273, -1.367969, -2.586083, -0.758337, 1.570796, 2.055069],accel_mss,speed_ms,0,blend_radius_m)
  movel([0.481001, -1.368865, -2.585468, -0.758056, 1.570796, 2.051797],accel_mss,speed_ms,0,blend_radius_m)
  movel([0.474434, -1.370965, -2.584022, -0.757402, 1.570796, 2.045231],accel_mss,speed_ms,0,blend_radius_m)
  movel([0.472989, -1.371456, -2.583683, -0.757250, 1.570796, 2.043785],accel_mss,speed_ms,0,blend_radius_m)
  movel([0.472799, -1.371633, -2.583560, -0.757195, 1.570796, 2.043595],accel_mss,speed_ms,0,blend_radius_m)
  movel([0.472675, -1.372000, -2.583307, -0.757082, 1.570796, 2.043471],accel_mss,speed_ms,0,blend_radius_m)
  movel([0.472651, -1.372400, -2.583030, -0.756959, 1.570796, 2.043448],accel_mss,speed_ms,0,blend_radius_m)
  speed_ms = 0.005
  movel([0.472651, -1.363527, -2.579005, -0.769857, 1.570796, 2.043448],accel_mss,speed_ms,0,blend_radius_m)
  speed_ms = 0.040
  movel([0.476821, -1.340541, -2.594336, -0.777512, 1.570796, 2.047618],accel_mss,speed_ms,0,blend_radius_m)
  speed_ms = 0.005
  movel([0.476821, -1.349572, -2.598463, -0.764353, 1.570796, 2.047618],accel_mss,speed_ms,0,blend_radius_m)
  speed_ms = 0.025
  movel([0.477677, -1.347959, -2.599526, -0.764904, 1.570796, 2.048473],accel_mss,speed_ms,0,blend_radius_m)
  movel([0.478294, -1.346339, -2.600590, -0.765460, 1.570796, 2.049091],accel_mss,speed_ms,0,blend_radius_m)
  movel([0.478658, -1.344752, -2.601629, -0.766008, 1.570796, 2.049454],accel_mss,speed_ms,0,blend_radius_m)
  movel([0.478760, -1.343233, -2.602620, -0.766537, 1.570796, 2.049556],accel_mss,speed_ms,0,blend_radius_m)
  movel([0.478382, -1.339736, -2.604888, -0.767764, 1.570796, 2.049178],accel_mss,speed_ms,0,blend_radius_m)
  movel([0.478408, -1.338690, -2.605564, -0.768135, 1.570796, 2.049205],accel_mss,speed_ms,0,blend_radius_m)
  movel([0.478593, -1.337680, -2.606215, -0.768494, 1.570796, 2.049389],accel_mss,speed_ms,0,blend_radius_m)
  movel([0.478986, -1.336760, -2.606806, -0.768823, 1.570796, 2.049782],accel_mss,speed_ms,0,blend_radius_m)
  movel([0.479645, -1.335982, -2.607306, -0.769101, 1.570796, 2.050441],accel_mss,speed_ms,0,blend_radius_m)
  movel([0.480625, -1.335334, -2.607721, -0.769334, 1.570796, 2.051421],accel_mss,speed_ms,0,blend_radius_m)
  movel([0.481492, -1.335098, -2.607872, -0.769419, 1.570796, 2.052289],accel_mss,speed_ms,0,blend_radius_m)
  movel([0.482252, -1.335197, -2.607809, -0.769383, 1.570796, 2.053048],accel_mss,speed_ms,0,blend_radius_m)
  movel([0.482905, -1.335552, -2.607581, -0.769256, 1.570796, 2.053701],accel_mss,speed_ms,0,blend_radius_m)
  movel([0.483890, -1.336704, -2.606842, -0.768843, 1.570796, 2.054687],accel_mss,speed_ms,0,blend_radius_m)
  movel([0.484469, -1.337923, -2.606058, -0.768408, 1.570796, 2.055265],accel_mss,speed_ms,0,blend_radius_m)
  movel([0.485197, -1.335855, -2.607387, -0.769147, 1.570796, 2.055994],accel_mss,speed_ms,0,blend_radius_m)
  movel([0.485588, -1.333878, -2.608652, -0.769859, 1.570796, 2.056384],accel_mss,speed_ms,0,blend_radius_m)
  movel([0.485773, -1.330063, -2.611077, -0.771248, 1.570796, 2.056569],accel_mss,speed_ms,0,blend_radius_m)
  movel([0.485880, -1.326195, -2.613517, -0.772677, 1.570796, 2.056677],accel_mss,speed_ms,0,blend_radius_m)
  movel([0.486175, -1.324147, -2.614800, -0.773442, 1.570796, 2.056971],accel_mss,speed_ms,0,blend_radius_m)
  movel([0.486781, -1.321976, -2.616155, -0.774258, 1.570796, 2.057577],accel_mss,speed_ms,0,blend_radius_m)
  movel([0.487335, -1.320582, -2.617021, -0.774786, 1.570796, 2.058131],accel_mss,speed_ms,0,blend_radius_m)
  movel([0.487908, -1.319452, -2.617721, -0.775216, 1.570796, 2.058704],accel_mss,speed_ms,0,blend_radius_m)
  movel([0.488491, -1.318572, -2.618266, -0.775552, 1.570796, 2.059287],accel_mss,speed_ms,0,blend_radius_m)
  movel([0.489074, -1.317931, -2.618661, -0.775797, 1.570796, 2.059870],accel_mss,speed_ms,0,blend_radius_m)
  movel([0.489642, -1.317515, -2.618918, -0.775956, 1.570796, 2.060439],accel_mss,speed_ms,0,blend_radius_m)
  movel([0.490193, -1.317306, -2.619047, -0.776037, 1.570796, 2.060989],accel_mss,speed_ms,0,blend_radius_m)
  movel([0.490709, -1.317289, -2.619057, -0.776043, 1.570796, 2.061506],accel_mss,speed_ms,0,blend_radius_m)
  movel([0.491186, -1.317453, -2.618956, -0.775980, 1.570796, 2.061982],accel_mss,speed_ms,0,blend_radius_m)
  movel([0.491611, -1.317781, -2.618753, -0.775854, 1.570796, 2.062408],accel_mss,speed_ms,0,blend_radius_m)
  movel([0.491974, -1.318257, -2.618460, -0.775672, 1.570796, 2.062770],accel_mss,speed_ms,0,blend_radius_m)
  movel([0.492480, -1.319590, -2.617636, -0.775163, 1.570796, 2.063276],accel_mss,speed_ms,0,blend_radius_m)
  movel([0.492629, -1.321327, -2.616558, -0.774504, 1.570796, 2.063426],accel_mss,speed_ms,0,blend_radius_m)
  movel([0.492348, -1.323346, -2.615301, -0.773742, 1.570796, 2.063144],accel_mss,speed_ms,0,blend_radius_m)
  movel([0.493591, -1.321653, -2.616356, -0.774380, 1.570796, 2.064387],accel_mss,speed_ms,0,blend_radius_m)
  movel([0.494597, -1.320010, -2.617376, -0.775003, 1.570796, 2.065393],accel_mss,speed_ms,0,blend_radius_m)
  movel([0.495417, -1.318404, -2.618369, -0.775616, 1.570796, 2.066213],accel_mss,speed_ms,0,blend_radius_m)
  movel([0.497377, -1.313599, -2.621321, -0.777469, 1.570796, 2.068173],accel_mss,speed_ms,0,blend_radius_m)
  movel([0.498859, -1.310219, -2.623380, -0.778791, 1.570796, 2.069655],accel_mss,speed_ms,0,blend_radius_m)
  movel([0.499616, -1.308827, -2.624223, -0.779339, 1.570796, 2.070412],accel_mss,speed_ms,0,blend_radius_m)
  movel([0.500393, -1.307640, -2.624940, -0.779809, 1.570796, 2.071190],accel_mss,speed_ms,0,blend_radius_m)
  movel([0.501171, -1.306658, -2.625532, -0.780199, 1.570796, 2.071967],accel_mss,speed_ms,0,blend_radius_m)
  movel([0.501934, -1.305878, -2.626001, -0.780510, 1.570796, 2.072731],accel_mss,speed_ms,0,blend_radius_m)
  movel([0.502667, -1.305294, -2.626352, -0.780743, 1.570796, 2.073464],accel_mss,speed_ms,0,blend_radius_m)
  movel([0.503355, -1.304905, -2.626585, -0.780899, 1.570796, 2.074152],accel_mss,speed_ms,0,blend_radius_m)
  movel([0.503982, -1.304707, -2.626704, -0.780978, 1.570796, 2.074779],accel_mss,speed_ms,0,blend_radius_m)
  movel([0.504532, -1.304696, -2.626710, -0.780982, 1.570796, 2.075329],accel_mss,speed_ms,0,blend_radius_m)
  movel([0.504990, -1.304870, -2.626606, -0.780913, 1.570796, 2.075786],accel_mss,speed_ms,0,blend_radius_m)
  movel([0.505340, -1.305221, -2.626395, -0.780772, 1.570796, 2.076136],accel_mss,speed_ms,0,blend_radius_m)
  movel([0.505569, -1.305747, -2.626080, -0.780562, 1.570796, 2.076366],accel_mss,speed_ms,0,blend_radius_m)
  movel([0.505661, -1.306444, -2.625660, -0.780284, 1.570796, 2.076458],accel_mss,speed_ms,0,blend_radius_m)
  movel([0.505600, -1.307307, -2.625140, -0.779941, 1.570796, 2.076396],accel_mss,speed_ms,0,blend_radius_m)
  movel([0.505372, -1.308332, -2.624522, -0.779535, 1.570796, 2.076168],accel_mss,speed_ms,0,blend_radius_m)
  movel([0.504963, -1.309512, -2.623808, -0.779069, 1.570796, 2.075759],accel_mss,speed_ms,0,blend_radius_m)
  movel([0.504361, -1.310843, -2.623001, -0.778545, 1.570796, 2.075158],accel_mss,speed_ms,0,blend_radius_m)
  movel([0.505882, -1.309678, -2.623708, -0.779003, 1.570796, 2.076678],accel_mss,speed_ms,0,blend_radius_m)
  movel([0.507291, -1.308414, -2.624472, -0.779502, 1.570796, 2.078088],accel_mss,speed_ms,0,blend_radius_m)
  movel([0.508613, -1.307071, -2.625283, -0.780035, 1.570796, 2.079409],accel_mss,speed_ms,0,blend_radius_m)
  movel([0.509871, -1.305667, -2.626128, -0.780594, 1.570796, 2.080667],accel_mss,speed_ms,0,blend_radius_m)
  movel([0.514730, -1.299885, -2.629580, -0.782925, 1.570796, 2.085526],accel_mss,speed_ms,0,blend_radius_m)
  movel([0.516568, -1.297775, -2.630828, -0.783786, 1.570796, 2.087364],accel_mss,speed_ms,0,blend_radius_m)
  movel([0.518895, -1.295391, -2.632232, -0.784766, 1.570796, 2.089692],accel_mss,speed_ms,0,blend_radius_m)
  movel([0.520143, -1.294383, -2.632824, -0.785183, 1.570796, 2.090940],accel_mss,speed_ms,0,blend_radius_m)
  movel([0.521391, -1.293655, -2.633250, -0.785484, 1.570796, 2.092187],accel_mss,speed_ms,0,blend_radius_m)
  movel([0.522003, -1.293434, -2.633379, -0.785576, 1.570796, 2.092800],accel_mss,speed_ms,0,blend_radius_m)
  movel([0.523177, -1.293343, -2.633433, -0.785614, 1.570796, 2.093973],accel_mss,speed_ms,0,blend_radius_m)
  movel([0.523727, -1.293507, -2.633336, -0.785546, 1.570796, 2.094523],accel_mss,speed_ms,0,blend_radius_m)
  movel([0.524119, -1.293909, -2.633101, -0.785379, 1.570796, 2.094915],accel_mss,speed_ms,0,blend_radius_m)
  movel([0.524203, -1.294537, -2.632733, -0.785119, 1.570796, 2.095000],accel_mss,speed_ms,0,blend_radius_m)
  movel([0.523804, -1.296075, -2.631830, -0.784484, 1.570796, 2.094600],accel_mss,speed_ms,0,blend_radius_m)
